(* IEC 61131-3 sources: IRIS-Project/LASAL CONTROL SOFTWARE/LasalProject_2025_09_12/Class/DiasMasterMain (part 3) *)

	push		  ecx
	push		  ebx

	L.eax		  (ebx+OneHandle.thisp)
	LZXW.ECX	(ebx+OneHandle.Address)
	push		  ecx
	push		  eax

	call		  CallUpdataRT
	add.esp		8

	pop			  ebx
	pop			  ecx

NextHandleRt
	add.ebx		sizeof (OneHandle)
	loop		  HandleLoopRt

LABEL_RtPostScan
//BLEERN START
  cmp.d     HwControl, 0
  jne       Rt_end

  call      UpdateRtPostScan_IM
//BLEERN ENDE

	jmp			  RT_end

// ****************************************************************
//  now we have to move the startpoint till we are 50usec before
// ****************************************************************

MovStartPoint

	//#SR001 Start
	L.EAX		  ud_DelayRealtime	//Time of Rt - Programm of IM
	CLR			  EDX
	L.ECX		  DmTmrResso*1000		// we have nanoseconds and we have to put in 25µs units
	DIV 		  ECX
	l.ebx		  eax
	//#SR001 End

	l.eax		  RtInterval

	sub.eax		ebx

	//#SR013 start
	cmp.b		  us_MuSecMode,1			//have we µs - Mode
	jne			  LABEL_Reserve_Std
	sub.eax		DmTimeReserveIM			//not so much reserve tim in µs - Mode
	jmp			  LABEL_EndReserve
LABEL_Reserve_Std
	//#SR013 end
	sub.eax		DmTimeReserveIM + 1		//ws005: just subtract 3 instead of ... (see above)			//#SR010 (make variable with define [instead of 3])
LABEL_EndReserve						//#SR013
  s.al		  (EDI+DmPllSyncDel)
	imul.ax		ax,DmTmrResso			//#SR009
	s.ax		  ui_RtStartPoint			//#SR009
	inc.b		  RtSSW					//ws005
	call		  LogRtSSW				//#SR008
	jmp			  RT_end

// ***********************************************************
//   read the calculated time
// ***********************************************************

ReadPoint
	clr			  eax
	l.al		  (edi+DmUserData)
	s.ax		  TimeBeforeNextSync
	inc.b		  RtSSW				//ws005
	call		  LogRtSSW			//#SR008
	jmp			  RT_end

// **********************************************************
//  now we are starting the RTProg
// **********************************************************

weAreSync
	call		  StartRealtimeProg
	inc.b		  RtSSW				//ws005
	call		  LogRtSSW			//#SR008
	jmp			  RT_end

// ***********************************************************
//   we have to wait that the PLL is locked before we start
// ***********************************************************
WaitForSync
	cmp.d		  release,16#FFFFFFFF
	je			  RT_end					// #fa 080103

	l			    (edi+DmPLLSyncState)
	test.al		DmPLLisLock
	jz			  WaitForSyncRet
	call		  StartRealtimeProg
	inc.b		  RtSSW				//ws005
	call		  LogRtSSW			//#SR008
	l.edi		  _IOSEGMENT			//#SR008
WaitForSyncRet
	L.AL		  (EDI+DmState)           // Start it always to keep the moduls alive
	OR.AL		  16#10
	S.AL		  (EDI+DmState)
	// #BS002

RT_end

	BT.W			StateCDiasSync+0,0
	JC				CDIASSyncOK
	L.EDI			CDIASSync // sync of CDIASBus
	L				  (EDI+2)
	S				  StateCDiasSync
CDIASSyncOK

	FC				WDCDIAS
RT_End1
	L.EAX	 		READY$UDINT

//#wp001
//============================ Profiler end======================================================
#ifdef  DiasMasterC_Profiler
	cmp.b 		DMC_Time_RT.initfl, 1				//schaun ob Delayzeit schon abgelaufen ist
	je			  LABEL_DMCEND
	pushad
	l.edi 		_LSL_POS
	l.edi 		( edi + DM_LSLPOS_SYSTIME )
	l.edi 		( edi + DM_LSLSYSTIME_MICROSEC )
	call		  edi								//OS_REadMicroSec - Funktion aufrufen
	s.eax 		DMC_Time_RT.stop					//Stopzeit speichern
	l.ebx 		DMC_Time_RT.start
	sub.eax		ebx								//Differenz berechnen
	sub.eax		DM_CPUconstant					//Zeit für OS_REadMicroSec - Funktion subtrahieren
	s.eax 		DMC_Time_RT.diff					//Ergebnis speicern
	l.ebx 		DMC_Time_RT.sum
	add.ebx 	eax								//Zur Summe addieren
	s.ebx 		DMC_Time_RT.sum					//Summe speichern
	l.ecx		  DMC_Time_RT.run
	inc 		  ecx								//Durchlaufzähler erhöhen
	s.ecx 		DMC_Time_RT.run					//Durchlaufzähler speichern
	cmp.eax		DMC_Time_RT._min					//mit Minimalzeit vergleichen
	jae			  LABEL_DMCcont
	s.eax 		DMC_Time_RT._min					//Minimalzeit speichern

LABEL_DMCcont
	cmp.eax 	DMC_Time_RT._max					//Mit Maximalzeit vergleichen
	jbe 		  LABEL_DMCcont1
	s.eax 		DMC_Time_RT._max					//Maximalzeit speichern

LABEL_DMCcont1
	l.eax		  ebx								//Summe in al laden
	imul.eax	eax,100							//*100 damit wir 2 Kommastellen haben
	x.edx 		edx
	idiv		  ecx								//durch Durchläufe dividieren
	s.eax		  DMC_Time_RT.avg					//Durchschnitt speichern
	popad

LABEL_DMCEND
	STI
#endif
//============================ Profiler end========================================================

END_FUNCTION
#endif

FUNCTION  DiasMasterMain::WDDIAS

	IF FirstModulFound <> 16#ff THEN	//ws005
	  IF DiasType <> 2 | RtSSw <> 4 THEN
 #IFNDEF MaxWatchdog	// #BS016
		IF ops.tAbsolute - timestamp$UDINT > 100ms | RtDebug = 1 THEN				//#SR011
			timestamp$UDINT := ops.tAbsolute;
 #ENDIF

			//**** Watchdog *************************************
			ReadKenn(FirstModulFound);

 #IFNDEF MaxWatchdog	// #BS016
		END_IF;
 #ENDIF
	  END_IF;
	END_IF;

	IF DiasType = 2 THEN
 #IFNDEF MaxWatchdog	// #BS016
		IF ops.tAbsolute - timestamp$UDINT > 100ms | RtDebug = 1 THEN				//#SR011
			timestamp$UDINT := ops.tAbsolute;
 #ENDIF

			IF (((_IOSegment$UDINT + DmControl)$^USINT)^ AND 2#10) = 0 & MasterON = 1 THEN
				MasterON := 0; // Risk is stopped => would be a watchdog
				IF Firstmodulfound <> 16#ff THEN		//ws005
          bdRTLogs.Bit6 := 1;
				END_IF;
				ImOff := 1;
			END_IF;

			//**** Watchdog for Risk (Xlinixversion 2.1) ****
			((_IOSegment$UDINT + DMWDRegister)$^USINT)^ := 1;

 #IFNDEF MaxWatchdog	// #BS016
		END_IF;
 #ENDIF
	END_IF;

END_FUNCTION

#ifdef _LSL_TARGETARCH_ARM
FUNCTION VIRTUAL GLOBAL DiasMasterMain::AddNOP
  VAR_INPUT
    RTCY		  : DINT;
    nCount		: DINT;
  END_VAR
  VAR
    i : DINT;
  END_VAR

  if (RTCY AND DmRealtime) = DmRealtime then
    ud_DelayRealtime += C_TimeNop;
  else
    ud_DelayCyclic += C_TimeNop;
  end_if;

  for i := 0 to (nCount-1) do
    (PtrCode + IPSub)^ := DbNop;

    IPSub += sizeof(RetStruct);
  end_for;

END_FUNCTION

#else
//
//	THR Aug. 21, 2003
//		Added function to add NOPs to the RISC program.  Unlike the
//		WAIT command, a NOP command CANNOT be interrupted by the
//		Cyclic Program.
//		Only for old DiasModuls
FUNCTION AWL VIRTUAL GLOBAL DiasMasterMain::AddNOP
  VAR_INPUT
    RTCY		  : DINT;
    nCount		: DINT;
  END_VAR

	l.eax		  RTCY
	and.eax		Dmrealtime

//#SR001 Start
	x.edx		  edx						//#SR003
	l.ebx		  nCount					//#SR003		//#SR009 (use ebx instead of eax register)
	imul.ebx	ebx,C_TimeNop			//#SR003		//#SR009
	CMP.EAX		Dmrealtime
	JNE			  LABEL_AN_NORT
	ADD.D		  ud_DelayRealtime,ebx	//#SR003		//#SR009
  JMP       LABEL_AN_TIMETAKEN
LABEL_AN_NORT
	ADD.D		  ud_DelayCyclic,ebx
//#SR001 End

LABEL_AN_TIMETAKEN

	call		  GetProgPointer

  l.ebx     PtrCode

	push		  ecx
	l.ecx		  nCount+0
an_loop
	l.b			  (edx+ebx),DbNop	   			// opcode NOP
	inc			  edx
	loop		  an_loop						//ws005: replaced dec,jnz with loop
	pop			  ecx

	l.eax		  RTCY
	and.eax		Dmrealtime
	call		  StoreNewPointers

END_FUNCTION
#endif

FUNCTION  DiasMasterMain::ErrorLocalSyncTrace

#ifdef HWC_LogError
  HWC_LogError(this, "@000A (DiasMasterMain::ErrorLocalSyncTrace) The constant 'NumberLocalSyncs' is defined too small !!! Remember: This is the number of maximum local Syncs !!!");
#else
	TRACE("The constant 'NumberLocalSyncs' is defined too small !!! Remember: This is the number of maximum local Syncs !!!");
#endif

END_FUNCTION

FUNCTION  DiasMasterMain::GetVerIMCIPC
  VAR_OUTPUT
    Ver(EAX)		: HDINT; // #BS016
  END_VAR
  VAR
    SigmaTekDevInfo : ^PCICONFDATA;
  END_VAR

#ifdef _LSL_TARGETARCH_X86
	SAVE_REG();
#endif

	IF pSPCIInfo <> NIL THEN
		SigmaTekDevInfo := SPCIINFO_FINDDEVICEBYNAME( "DIASIM" , 0 );
		Ver := 0;
		IF SigmaTekDevInfo <> NIL THEN
			Ver$USINT := SigmaTekDevInfo^.Version;
		END_IF;
	ELSE
		Ver := 0; // Error in OS - Interface (shouldn't be)
	END_IF;

#ifdef _LSL_TARGETARCH_X86
	RESTORE_REG();
#endif

(*
other funktions:

VAR
	pSPCIInfo     	: ^LSL_SPCIINFO;
	SigmatTekDevs	: DINT;
	SigmaTekDevInfo : ^PCICONFDATA;
	Version : USINT;
	Index : DINT;
	BaseAddress : ^VOID;
	BaseAddressLEN : UDINT;
END_VAR

	if OS_CILGET("PCICONFIG", #pSPCIInfo) then
		state:= 1;
	else
		state:= 0;
	end_if;

	// Anzahl der Einträge im InfoBlock
	SigmatTekDevs := SPCIINFO_GETDEVICECOUNT();

	for Index := 0 to SigmatTekDevs-1 do
		SigmaTekDevInfo := SPCIINFO_GETDEVICEBYINDEX( Index );
		Version := SigmaTekDevInfo^.Version;
	end_for;

	// z.B. PLL
	SigmaTekDevInfo := SPCIINFO_FINDDEVICEBYNAME( "PLL", 0 );
	SigmaTekDevInfo := SPCIINFO_FINDDEVICE( 16#0E08, 0 );
	BaseAddress := SPCIINFO_GETADDRESS( SigmaTekDevInfo );
	BaseAddressLen := SPCIINFO_GETADDRESSLEN( SigmaTekDevInfo );

	// z.B. CDIAS
	SigmaTekDevInfo := SPCIINFO_FINDDEVICEBYNAME( "CDiasBus", 0 );
	SigmaTekDevInfo := SPCIINFO_FINDDEVICE( 16#0500, 0 );
	BaseAddress := SPCIINFO_GETADDRESS( SigmaTekDevInfo );
	BaseAddressLen := SPCIINFO_GETADDRESSLEN( SigmaTekDevInfo );

*)

END_FUNCTION

FUNCTION DiasMasterMain::TraceAsyncError
	VAR_INPUT
		Place 	: UDINT;(* := 255 *)
	END_VAR
  VAR
    ptr		  : ^USINT;
    tracewd	: USINT;		// #BS012
    LogStr  : ARRAY [0..255] OF CHAR;
    NumStr  : ARRAY [0..9] OF CHAR;
  END_VAR

	if ( MasterOn <> 0 ) then		//#SR016	( because otherwise we have a lot of event messages

#ifdef _LSL_TARGETARCH_X86
		SAVE_REG();
#endif
		// #BS012 Start
		tracewd := 0;
		IF CDIASType = 2 THEN // CIPC
			IF ((CDiasI2CWatchdog+2)^ AND 1) = 1 THEN // watchdogstatus (Bit0 = 1 => watchdog)
#ifdef HWC_LogError
        HWC_LogError(this, "@0578 (DiasMasterMain::TraceAsyncError) Watchdog on CDIAS and DIAS - Bus occured !! (The RtTask of DiasMasterC - Class was set Off for more than 30ms => Hardwarereset on DIAS and CDIAS - Bus)");
#else
				// Watchdog on CDIAS and DIAS - Bus occured !! (The RtTask of DiasMasterC - Class was set Off for more than 30ms => Hardwarereset on DIAS and CDIAS - Bus)
				Trace("DiasMaster: Watchdog on CDIAS and DIAS - Bus occured !! (The RtTask of DiasMasterC - Class was set Off for more than 30ms => Hardwarereset on DIAS and CDIAS - Bus)");
				//#SR008 start
				if p_KernelLog <> NIL then
					OS_KernelLog0( "DiasMaster: Watchdog on CDIAS and DIAS - Bus occured !! (The RtTask of DiasMasterC - Class was set Off for more than 30ms => Hardwarereset on DIAS and CDIAS - Bus)" );
				end_if;
				//#SR008 end
#endif
			ELSE
				tracewd := 1;
			END_IF;
		END_IF;
		// #BS012 End
		ptr$UDINT := _IOSegment$UDINT + DMControl;
		ptr^ := 1; // Chip on risk off
		ImOff := 1;
		MasterOn := 0;
#ifdef HWC_LogError
    HWC_LogError(this, "@0582 (DiasMasterMain::TraceAsyncError) Timeout on asynchron methods !! => DiasBus is set off!!");
#else
		TRACE("DiasMaster: Timeout on asynchron methods !! => DiasBus is set off!!");
		//#SR008 start
		if p_KernelLog <> NIL then
			OS_KernelLog0( "DiasMaster: Timeout on asynchron methods !! => DiasBus is set off!!" );
		end_if;
#endif

#ifndef DIASMASTER_DISABLE_DIAS_ERROR_ON_DIRECT_ACCESS
    // if we got a place => create a dias error
    if Place <> 255 then

#ifdef HWC_LogValue1
      HWC_LogValue1(this, "@05F0 (DiasMasterMain::TraceAsyncError) Dias Error occured at place 0x{0}", Place);
#else
      _strcpy(dest:=#LogStr[0], src:="(DiasMasterMain::TraceAsyncError) Dias Error occured at place 0x");
      _itoa(udNumber:=Place, pString:=#NumStr[0]);
      _strcat(dest:=#LogStr[0], src:=#NumStr[0]);
      TRACE(#LogStr[0]);
      if p_KernelLog <> NIL then
        OS_KernelLog0(#LogStr[0]);
      end_if;
#endif

      _strcpy(dest:=#LogStr[0], src:="exec climsg 25 Dias Error occured at place 0x");
      _itoa(udNumber:=Place, pString:=#NumStr[0]);
      _strcat(dest:=#LogStr[0], src:=#NumStr[0]);

      To_OSKernel.AddToServiceProvider(command:=#LogStr[0], immediatly:=1);
    end_if;
#endif

		//#SR008 end
		// #BS012 Start
		IF tracewd THEN
#ifdef HWC_LogError
      HWC_LogError(this, "@058C (DiasMasterMain::TraceAsyncError) But no Watchdog on CDIAS and DIAS - Bus");
#else
			Trace("DiasMaster: But no Watchdog on CDIAS and DIAS - Bus");
			//#SR008 start
			if p_KernelLog <> NIL then
				OS_KernelLog0( "DiasMaster: But no Watchdog on CDIAS and DIAS - Bus" );
			end_if;
			//#SR008 end
#endif
		END_IF;
		// #BS012 End
#ifdef _LSL_TARGETARCH_X86
		RESTORE_REG();
#endif
	end_if;						//#SR016

END_FUNCTION

FUNCTION  DiasMasterMain::GetMuSec
  VAR_OUTPUT
    value(EAX)		: UDINT;
  END_VAR

#ifdef _LSL_TARGETARCH_X86
	SAVE_REG();
#endif
	value := OS_ReadMicroSec();

#ifdef _LSL_TARGETARCH_X86
	RESTORE_REG();
#endif

END_FUNCTION

#ifdef _LSL_TARGETARCH_ARM
FUNCTION VIRTUAL GLOBAL DiasMasterMain::AddRdKenn
  VAR_INPUT
    Adress		: HSINT;
    RTCY		: DINT;
    thisp		: ^void;
    callOptions 	: USINT;
  END_VAR
  VAR_OUTPUT
    Handle		: DINT;
  END_VAR

  if (RTCY AND DmRealtime) = DmRealtime then
    ud_DelayRealtime += C_TimeReadKennung;
    ui_RtDIASAccesses += 1;
  else
    ud_DelayCyclic += C_TimeReadKennung;
    ui_CyDIASAccesses += 1;
  end_if;

  (PtrCode + IPSub + RdKennStruct.Opc)^   := DbRdKenn;
  (PtrCode + IPSub + RdKennStruct.ModAdr)^ := Adress;

  ARM_EAX := RTCY$UDINT;
  ARM_EDI := thisp$UDINT;
  GetHandle(RdKennStruct.Data, callOptions);
  Handle := ARM_EAX$DINT;
  IPSub += sizeof(RdKennStruct);

END_FUNCTION

#else
// to read the identifier of a modul

FUNCTION AWL VIRTUAL GLOBAL DiasMasterMain::AddRdKenn
	VAR_INPUT
		Adress 	: HSINT;
		RTCY 	: DINT;
		thisp 	: ^void;
		callOptions 	: USINT;
	END_VAR
	VAR_OUTPUT
		Handle 	: DINT;
	END_VAR

	l.eax		  RTCY
	and.eax		Dmrealtime

//#SR001 Start
	CMP.EAX		Dmrealtime
	JNE			  LABEL_ARK_NORT
	ADD.D		  ud_DelayRealtime,C_TimeReadKennung
	inc.w		  ui_RtDIASAccesses			//#SR021
  JMP       LABEL_ARK_TIMETAKEN

LABEL_ARK_NORT
	ADD.D		  ud_DelayCyclic,C_TimeReadKennung
	inc.w		  ui_CyDIASAccesses
//#SR001 End

LABEL_ARK_TIMETAKEN

	call		  GetProgPointer

  l.ebx     PtrCode

	l.b			  (edx+ebx+RdKennStruct.Opc),DbRdKenn	   			// opcode read identifier
	l			    Adress					// adress of dias modul
	s			    (edx+ebx+RdKennStruct.ModAdr)

	l.ax		  RTCY+0
	l.edi		  thisp				    // to put into then handle

  push.b    callOptions

	push.d		RdKennStruct.Data			// direct pointer on the data
	call		  GetHandle
  add.esp   5

	s.eax		  Handle
	add.edx		sizeof (RdKennStruct)

	l.eax		  RTCY
	and.eax		Dmrealtime
	call		  StoreNewPointers

END_FUNCTION
#endif

#ifdef _LSL_TARGETARCH_ARM
FUNCTION VIRTUAL GLOBAL DiasMasterMain::AddMove
  VAR_INPUT
    RTCY		: DINT;
    thisp		: ^void;
    callOptions 	: USINT;
    SourceAddr 	: HDINT;
    DestAddr 	: HDINT;
    MoveLen 	: UDINT;
    pEnable 	: ^USINT;
    Settings 	: HDINT;
  END_VAR
  VAR_OUTPUT
    HandleMove		: DINT;
  END_VAR

  if (RTCY AND DmRealtime) = DmRealtime then
    ud_DelayRealtime += C_TimeMove;
  else
    ud_DelayCyclic += C_TimeMove;
  end_if;

  (PtrCode + IPSub + MoveStruct.Opc)^               := DbMov;
  (PtrCode$^HINT + IPSub + MoveStruct.Source)^      := (IPSub + MoveStruct.Destination)$HINT;
  (PtrCode$^HINT + IPSub + MoveStruct.Destination)^ := (IPSub + MoveStruct.Destination)$HINT;

  ARM_EAX := RTCY$UDINT;
  ARM_EDI := thisp$UDINT;
  GetHandle(MoveStruct.Source, callOptions);
  HandleMove := ARM_EAX$DINT;
  IPSub += sizeof(MoveStruct);

END_FUNCTION

#else
// BS 14.11.2001
// This command is to switch for example a bank back in im routine.
//
//[#ENGLISH]
//[<HandleMove]pointer on source (2 Byte further is destination)

FUNCTION AWL VIRTUAL GLOBAL DiasMasterMain::AddMove
	VAR_INPUT
		RTCY 	: DINT;
		thisp 	: ^void;
		callOptions 	: USINT;
		SourceAddr 	: HDINT;
		DestAddr 	: HDINT;
		MoveLen 	: UDINT;
		pEnable 	: ^USINT;
		Settings 	: HDINT;
	END_VAR
	VAR_OUTPUT
		HandleMove 	: DINT;
	END_VAR

	l.eax		  RTCY
	and.eax		Dmrealtime

//#SR001 Start
	CMP.EAX		Dmrealtime
	JNE			  LABEL_AM_NORT
	ADD.D		  ud_DelayRealtime,C_TimeMove
  JMP       LABEL_AM_TIMETAKEN

LABEL_AM_NORT
  ADD.D		  ud_DelayCyclic,C_TimeMove
//#SR001 End

LABEL_AM_TIMETAKEN

	call		  GetProgPointer

  l.ebx     PtrCode

	l.b			  (edx+ebx+MoveStruct.Opc),DbMov	   			// opcode read identifier

	L.EAX		  EDX
	ADD.EAX		MoveStruct.Destination
	S.AX		  (edx+ebx+MoveStruct.Source) // read destination
	S.AX		  (edx+ebx+MoveStruct.Destination) // save on destination

	l.ax		  RTCY+0
	l.edi		  thisp				    // to put into then handle

  push.b    callOptions

	push.d		MoveStruct.Source			// direct pointer on the data
	call		  GetHandle
  add.esp 5

	s.eax		  HandleMove
	add.edx		sizeof (MoveStruct)

	l.eax		  RTCY
	and.eax		Dmrealtime
	call		  StoreNewPointers

END_FUNCTION
#endif

FUNCTION VIRTUAL GLOBAL DiasMasterMain::GetCDiasPlaceIoSegment
  VAR_INPUT
    place		: UDINT;
  END_VAR
  VAR_OUTPUT
    IOSegment		: ^USINT;
  END_VAR

	IOSegment$UDINT :=  CDiasHwPointer$UDINT + (place*16#100)$UDINT;

END_FUNCTION

//[#ENGLISH]
//[<StateSync]0 = Busy | 1 = Sync | 2 = TimeOut
#ifdef _LSL_TARGETARCH_ARM
FUNCTION DiasMasterMain::CheckSyncModules
  VAR_INPUT
    TimeStampStart		: UDINT;
  END_VAR
  VAR_OUTPUT
    StateSync		: UDINT;
  END_VAR
  VAR
    pModule : ^WaitSyncCall;
    i : UDINT;
    MaxTime : UDINT;
  END_VAR

  // init with synchron
  StateSync := 1;

  // check if there are any sync calls
  if DiasSync.NumberCalls then
    pModule := #DiasSync.Modules[0];
    MaxTime := 0;

    // search for the max possible sync time
    for i := 0 to (DiasSync.NumberCalls - 1) do
      if (pModule^.SyncState = 0) & (pModule^.WaitTime > MaxTime) then
        MaxTime := pModule^.WaitTime;   // save the maxtime
      end_if;

      pModule += sizeof(WaitSyncCall);
    end_for;
    DiasSync.ActMaxTime := MaxTime;

    pModule := #DiasSync.Modules[0];

    // search if modules are ready
    for i := 0 to (DiasSync.NumberCalls - 1) do
      if (pModule^.SyncState = 0) then
        pModule^.SyncState := CallGetSync(thisp:=pModule^.thisp);
        if pModule^.SyncState = 0 then
          StateSync := 0;   // busy
        end_if;
      end_if;

      pModule += sizeof(WaitSyncCall);
    end_for;

    if (StateSync = 0) & ((ops.tAbsolute - TimeStampStart) > DiasSync.ActMaxTime) then
      StateSync := 2;   // timeout
    end_if;
  end_if;

END_FUNCTION
#else
FUNCTION AWL DiasMasterMain::CheckSyncModules
  VAR_INPUT
    TimeStampStart		: UDINT;
  END_VAR
  VAR_OUTPUT
    StateSync		: UDINT;
  END_VAR

// #BS014 Start
// init with synchron
	L.D			  StateSync,1

// check if there are any sync calls
	L.ECX		  DiasSync.NumberCalls
	JECXZ		  SyncReady

// search for the max possible sync time
	L.EDI		  #DiasSync.Modules[0]
	X.EAX		  EAX
SearchTime
	CMP.B		  (EDI+WaitSyncCall.SyncState),1	// if the modul is sync we cancel it
	JE			  NextObjectTime
	CMP.EAX		(EDI+WaitSyncCall.WaitTime)
	JAE			  NextObjectTime
	L.EAX		  (EDI+WaitSyncCall.WaitTime)		// save the maxtime
NextObjectTime
	ADD.EDI		SIZEOF(WaitSyncCall)
	LOOP		  SearchTime

	S.EAX		  DiasSync.ActMaxTime

// search if modules are ready
	L.EDI		  #DiasSync.Modules[0]
	L.ECX		  DiasSync.NumberCalls

SyncSearch

	CMP.B		  (EDI+WaitSyncCall.SyncState),1
	JE			  NextObject

	PUSH		  EDI
	PUSH		  ESI
	PUSH		  ECX

	X.AL		  AL

	L.EDI		  (EDI+WaitSyncCall.thisp)
	CALL		  CallGetSync

	POP			  ECX
	POP			  ESI
	POP			  EDI

	S.AL		  (EDI+WaitSyncCall.SyncState)
	CMP.AL	  1	// if sync then next obj
	JE			  NextObject
	L.D			  StateSync,0 // busy
NextObject
	ADD.EDI		SIZEOF(WaitSyncCall)
	LOOP		  SyncSearch

	CMP.D		  StateSync,1
	JE			  SyncReady

	L.EAX		  ops.tAbsolute
	SUB.EAX		TimeStampStart
	CMP.EAX		DiasSync.ActMaxTime
	JBE			  EndSyncCheck

	L.D			  StateSync,2 // timeout
	JMP			  EndSyncCheck

SyncReady

EndSyncCheck
// #BS014 End

END_FUNCTION
#endif

FUNCTION  DiasMasterMain::CallGetSync
  VAR_INPUT
    thisp(EDI)		: pHwBase;
  END_VAR
  VAR_OUTPUT
    syncchron(AL)		: USINT;
  END_VAR

	syncchron := thisp^.CheckSync();

END_FUNCTION

FUNCTION VIRTUAL GLOBAL DiasMasterMain::AddWaitSync
  VAR_INPUT
    thisp		: pVoid;
    MaxWaitTime		: UDINT;
  END_VAR

	IF DiasSync.NumberCalls * SIZEOF(WaitSyncCall) < SIZEOF(DiasSync.Modules) THEN
		DiasSync.Modules[DiasSync.NumberCalls$SINT].thisp$pVoid 	:= thisp;// #BS016
		DiasSync.Modules[DiasSync.NumberCalls$SINT].WaitTime := MaxWaitTime;// #BS016
		DiasSync.NumberCalls += 1;

		IF MaxWaitTime > DiasSync.ActMaxTime THEN
			DiasSync.ActMaxTime	:= MaxWaitTime;
		END_IF;
	ELSE

#ifdef HWC_LogError
    HWC_LogError(this, "@000B (DiasMasterMain::AddWaitSync) The constant 'MaxSyncModules' is defined too small !!!");
#else
		TRACE("The constant 'MaxSyncModules' is defined too small !!!");
#endif
	END_IF;

END_FUNCTION

FUNCTION VIRTUAL GLOBAL DiasMasterMain::Release::Read
	VAR_OUTPUT
		output (EAX) 	: HDINT;
	END_VAR

	output := Release;

END_FUNCTION

FUNCTION VIRTUAL GLOBAL DiasMasterMain::Chipstate::Read
  VAR_OUTPUT
    output		: DINT;
  END_VAR

	output := Chipstate;

END_FUNCTION

FUNCTION VIRTUAL GLOBAL DiasMasterMain::RiscState::Read
  VAR_OUTPUT
    output		: DINT;
  END_VAR

	output := RiscState;

END_FUNCTION

FUNCTION VIRTUAL GLOBAL DiasMasterMain::TimeAtRtPreEnd::Read
  VAR_OUTPUT
    output		: DINT;
  END_VAR

	output := TimeAtRtPreEnd;

END_FUNCTION

FUNCTION VIRTUAL GLOBAL DiasMasterMain::DIASRetryCounter::Read
  VAR_OUTPUT
    output		: DINT;
  END_VAR

	output := DIASRetryCounter;

END_FUNCTION

FUNCTION VIRTUAL GLOBAL DiasMasterMain::MasterON::Read
  VAR_OUTPUT
    output		: DINT;
  END_VAR

	output := MasterON;

END_FUNCTION

FUNCTION  DiasMasterMain::Risc_Off

#ifdef HWC_LogError
  HWC_LogError(this, "@0596 (DiasMasterMain::Risc_Off) RISC is set of -> DiasMasterOn = 0 and ImOff = 1");
#else
	TRACE("DiasMaster: RISC is set of -> DiasMasterOn = 0 and ImOff = 1");
	//#SR008 start
	if p_KernelLog <> NIL then
		OS_KernelLog0( "DiasMaster: RISC is set of -> DiasMasterOn = 0 and ImOff = 1" );
	end_if;
	//#SR008 end
#endif
	ImOff := 1;
	MasterOn := 0;

END_FUNCTION

#ifdef _LSL_TARGETARCH_ARM
FUNCTION VIRTUAL GLOBAL DiasMasterMain::AddIRQScan
  VAR_INPUT
    Place		: USINT;
    RTCY		: DINT;
    thisp		: ^void;
    callOptions 	: USINT;
  END_VAR
  VAR_OUTPUT
    Handle		: DINT;
  END_VAR

  if (RTCY AND DmRealtime) = DmRealtime then
    ud_DelayRealtime += C_TimeIRQScan;
  else
    ud_DelayCyclic += C_TimeIRQScan;
  end_if;

  (PtrCode + IPSub + IRQScanStruct.Opc)^    := DbIRQScan;
  (PtrCode + IPSub + IRQScanStruct.ModAdr)^ := Place;

  ARM_EAX := RTCY$UDINT;
  ARM_EDI := thisp$UDINT;
  GetHandle(IRQScanStruct.Data, callOptions);
  Handle := ARM_EAX$DINT;
  IPSub += sizeof(IRQScanStruct);

END_FUNCTION

#else
//[#ENGLISH]
//[>Place]modul number
FUNCTION AWL VIRTUAL GLOBAL DiasMasterMain::AddIRQScan
	VAR_INPUT
		Place 	: USINT;
		RTCY 	: DINT;
		thisp 	: ^void;
		callOptions 	: USINT;
	END_VAR
	VAR_OUTPUT
		Handle 	: DINT;
	END_VAR

	l.eax		  RTCY
	and.eax		Dmrealtime

	CMP.EAX		Dmrealtime
	JNE			  LABEL_AIRQ_NORT
	ADD.D		  ud_DelayRealtime,C_TimeIRQScan
  JMP       LABEL_AIRQ_TIMETAKEN

LABEL_AIRQ_NORT
	ADD.D		  ud_DelayCyclic,C_TimeIRQScan

LABEL_AIRQ_TIMETAKEN

	call		  GetProgPointer

  l.ebx     PtrCode

	l.b			  (edx+ebx+IRQScanStruct.Opc),DbIRQScan	   			// opcode IRQ identifier
	l			    Place					// place of dias modul
	s			    (edx+ebx+IRQScanStruct.ModAdr)

	l.ax		  RTCY+0
	l.edi		  thisp				    // to put into then handle

  push.b    callOptions

	push.d		IRQScanStruct.Data			// direct pointer on the data
	call		  GetHandle
  add.esp   5

	s.eax		  Handle
	add.edx		sizeof (IRQScanStruct)

	l.eax		  RTCY
	and.eax		Dmrealtime
	call		  StoreNewPointers

END_FUNCTION
#endif

#ifdef _LSL_TARGETARCH_ARM
FUNCTION VIRTUAL GLOBAL DiasMasterMain::IRQScan
  VAR_INPUT
    Place		: udint;
  END_VAR
  VAR_OUTPUT
    Data		: DINT;
  END_VAR
  VAR
    Time1, Time2  : UDINT;
    TimeoutFlag   : DINT;
  END_VAR

  if (DiasType = 2) & (ImOff = FALSE) then
#ifdef _LSL_TARGETARCH_X86
    Save_Flg();
    CLI();          // needed for async read
#endif

    Time1 := Time2 := OS_ReadMicroSec();

    while ((Time2 - Time1) <= DmConstTimeOut) do
      Time2 := OS_ReadMicroSec()
      if (_IOSegment$^USINT + DmCmdBuf1)^ AND 1 then
        exit;
      end_if;
    end_while;

    (_IOSegment$^USINT+1+DmCmdBuf1+IRQScanStruct.ModAdr)^ := Place$USINT;
    (_IOSegment$^USINT + DmCmdBuf1)^ := 0; // kill ready
    (_IOSegment$^USINT+1+DmCmdBuf1+IRQScanStruct.Opc)^ := DbIRQScan;

    Time1 := Time2 := OS_ReadMicroSec();
    TimeoutFlag := 1;

    while ((Time2 - Time1) <= DmConstTimeOut) do
      Time2 := OS_ReadMicroSec()
      if (_IOSegment$^USINT + DmCmdBuf1)^ AND 1 then
        Data := to_dint((_IOSegment$^USINT+1+DmCmdBuf1+IRQScanStruct.Data)^);
        TimeoutFlag := 0;
        exit;
      end_if;
    end_while;

    if TimeoutFlag then
      // timeout
      TraceAsyncError();
      Data := 0;
    end_if;

#ifdef _LSL_TARGETARCH_X86
    Restore_Flg();
#endif
  end_if;

END_FUNCTION

#else

FUNCTION AWL VIRTUAL GLOBAL DiasMasterMain::IRQScan
  VAR_INPUT
    Place		: udint;
  END_VAR
  VAR_OUTPUT
    Data		: DINT;
  END_VAR

  //ws005: moved to the start, since these cmp are critical
	cmp.b		  DiasType,2		//ws005
	jne			  LABEL_End		// --> it is a new Master

  CMP.B		  ImOff,1
	JE			  LABEL_End
  // /ws005

	push		  edi
	push		  ebx
	push		  eax

	L.EDI		  _IOSEGMENT

	CLR 		  EAX

 	L.ebx		  Place

	PUSHF
	CLI // needed for async read

	FC			  GetMuSec
	S.EAX		  EDX
BSyIRQ
	FC			  GetMuSec
	SUB.EAX		EDX
	TST.B		  (EDI+DmCmdBuf1),1
	JNZ			  BSyIRQConti
	CMP.EAX		DmConstTimeOut
	JA			  TimeOutError
	JMP			  BSyIRQ
BSyIRQConti

	S.Bl		  (EDI+1+DmCmdBuf1+IRQScanStruct.ModAdr)
	L.b			  (EDI+DmCmdBuf1),0		// Ready Töten
	L.B			  (EDI+1+DmCmdBuf1+IRQScanStruct.Opc),DbIRQScan

	FC			  GetMuSec
	S.EAX		  EDX
NixDaIRQ
	FC			  GetMuSec
	SUB.EAX		EDX
	TST.B		  (EDI+DmCmdBuf1),1
	JNZ			  IRQScanOkIM
	CMP.EAX		DmConstTimeOut
	JA			  TimeOutError
	JMP			  NixDaIRQ

TimeOutError
	POPF
  L.EAX     Place
  PUSH      EAX
	FC			  TraceAsyncError
  ADD.ESP   4
	L.D			  Data,0
	JMP			  LABEL_End1  //ws005

IRQScanOkIM
	LZXB.EAX	(EDI+1+DmCmdBuf1+IRQScanStruct.Data)
//	POPF				//#SR017
	S.EAX		  Data

LABEL_End1    //ws005
	POPF				//#SR017
	pop			  eax
	pop			  ebx
	pop			  edi

LABEL_End     //ws005

END_FUNCTION
#endif

//[#ENGLISH]
// This function updates the DIAS retry counter (using a function provided by the OS)
// [Globals]	_LSL_POS			:R		:OS interface structure
// [Members]	oldErrorCounter		:R/W	:calculate change
//			(S)	DiasRetryCounter	:W		:update retry counter
// [Locals]		us_actcount			:R/W	:currently read value
//				di_oldcount			:R/W	:temporary storeage of the previous value
FUNCTION DiasMasterMain::UpdateRetryCounter
  VAR
    us_actcount : usint;
    di_oldcount : dint;
    di_ret	    : dint;		//ws005
  END_VAR;

	if( pDIAS <> NIL )then	// CPU has a DIAS bus (for now only valid for CCL081)
		//ws005: consider the return value
		di_ret := OS_DIAS_ReadRegister( pDIAS, ( DIASRetryCounterOffset + 0 )$uint,  #us_actcount );
    di_oldcount := oldErrorCounter;
    oldErrorCounter := to_dint( us_actcount );
    DiasRetryCounter += oldErrorCounter - di_oldcount;
	end_if;

END_FUNCTION

//[#ENGLISH]
//Function gives back the Dias Adress, of the module which
//answer to the global sync.
FUNCTION VIRTUAL GLOBAL DiasMasterMain::GetSyncModuleNumber
  VAR_OUTPUT
    us_ModuleNr		: USINT;
  END_VAR

	us_ModuleNr := us_SyncModule;

END_FUNCTION

//[#ENGLISH]
//Function for logging Realtime steps at startup
FUNCTION  DiasMasterMain::LogRtSSW

  case RtSSW of

    1:		bdRTLogs.Bit1 := 1; //OS_KernelLog0( "DiasMaster: Pll is locked and Rt programm of intelligent master starts (1)"); 	//#SR021

    2:		bdRTLogs.Bit2 := 1; //OS_KernelLog1( "DiasMaster: We are Sync -> Rt programm of intelligent master starts again (Sync Module Place: %d) (2)", us_SyncModule ); 		//#SR021

    3:		bdRTLogs.Bit3 := 1; //OS_KernelLog2( "DiasMaster: MoveStartPointer -> Start moment of IM - programm is set (Rt - Startpoint: %dus, AddTime: %dns) (3)", ui_RtStartpoint, ui_AddTime );	//#SR021

    4:		bdRTLogs.Bit4 := 1; //OS_KernelLog1( "DiasMaster: One Time point was read -> start updating realtime tasks now (%d Rt - Dias accesses) (4)", ui_RtDIASAccesses );			//#SR021

  end_case;

END_FUNCTION

FUNCTION  DiasMasterMain::WriteRTLogs

  if bdRTLogs then
    if p_KernelLog <> NIL then
      if bdRTLogs.Bit1 then
        bdRTLogs.Bit1 := 0;
#ifdef HWC_LogError
        HWC_LogError(this, "@0514 (DiasMasterMain::WriteRTLogs) Pll is locked and Rt programm of intelligent master starts (1)");
#else
        if p_KernelLog <> NIL then
          OS_KernelLog0( "DiasMaster: Pll is locked and Rt programm of intelligent master starts (1)"); 	//#SR021
        end_if;
#endif
      end_if;
      if bdRTLogs.Bit2 then
        bdRTLogs.Bit2 := 0;
#ifdef HWC_LogValue1
        HWC_LogValue1(this, "@051E (DiasMasterMain::WriteRTLogs) We are Sync -> Rt programm of intelligent master starts again (Sync Module Place: {0}) (2)", us_SyncModule);
#else
        if p_KernelLog <> NIL then
          OS_KernelLog1( "DiasMaster: We are Sync -> Rt programm of intelligent master starts again (Sync Module Place: %d) (2)", us_SyncModule ); 		//#SR021
        end_if;
#endif
      end_if;
      if bdRTLogs.Bit3 then
        bdRTLogs.Bit3 := 0;
#ifdef HWC_LogValue2
        HWC_LogValue2(this, "@0528 (DiasMasterMain::WriteRTLogs) MoveStartPointer -> Start moment of IM - programm is set (Rt - Startpoint: {0}us, AddTime: {1}ns) (3)", ui_RtStartpoint, ui_AddTime);
#else
        if p_KernelLog <> NIL then
          OS_KernelLog2( "DiasMaster: MoveStartPointer -> Start moment of IM - programm is set (Rt - Startpoint: %dus, AddTime: %dns) (3)", ui_RtStartpoint, ui_AddTime );	//#SR021
        end_if;
#endif
      end_if;
      if bdRTLogs.Bit4 then
        bdRTLogs.Bit4 := 0;
#ifdef HWC_LogValue1
        HWC_LogValue1(this, "@0532 (DiasMasterMain::WriteRTLogs) One Time point was read -> start updating realtime tasks now (%d Rt - Dias accesses) (4)", ui_RtDIASAccesses);
#else
        if p_KernelLog <> NIL then
          OS_KernelLog1( "DiasMaster: One Time point was read -> start updating realtime tasks now (%d Rt - Dias accesses) (4)", ui_RtDIASAccesses );			//#SR021
        end_if;
#endif
      end_if;
    end_if;
  end_if;

  //Trace Message for Timesliceerror
	if us_FirstTimeSliceStart = 1 (* //#SR017 & ud_ErrorCountTimeSliceStart >= 10*) then

		us_FirstTimeSliceStart := 2;
#ifdef HWC_LogError
    HWC_LogError(this, "@05A0 (DiasMasterMain::Trace_JitterError) [SL] Rt of IM starts while Rt of DiasMaster is running!!");
#else
		trace("DiasMaster: Rt of IM starts while Rt of DiasMaster is running!!");
		if p_KernelLog <> NIL then
			OS_KernelLog0( "DiasMaster: Rt of IM starts while Rt of DiasMaster is running!!" );
		end_if;
#endif

	elsif us_FirstTimeSliceEnd = 1 (* //#SR017 & ud_ErrorCountTimeSliceEnd >= 10*) then

		us_FirstTimeSliceEnd := 2;
#ifdef HWC_LogError
    HWC_LogError(this, "@05AA (DiasMasterMain::Trace_JitterError) [SL] Timeslice overrun!!");
#else
		trace("DiasMaster: Timeslice overrun!!");
		if p_KernelLog <> NIL then
			OS_KernelLog0( "DiasMaster: Timeslice overrun!!" );
		end_if;
#endif
	end_if;

  //Watchdog Error CDIAS
  if bdRTLogs.Bit5 then
    if RTSSW <> 4 then
#ifdef HWC_LogError
      HWC_LogError(this, "@0564 (DiasMasterMain::WdCDIAS) Watchdog Error (RTSSW<>4) -> DiasMasterOn = 0 and ImOff = 1");
#else
      // Watchdog on CDIAS and DIAS - Bus occured !! (The RtTask of DiasMasterC - Class was set Off for more than 30ms => Hardwarereset on DIAS and CDIAS - Bus)
      Trace("Watchdog Error (RTSSW<>4) -> DiasMasterOn = 0 and ImOff = 1");
      //#SR008 start
      if p_KernelLog <> NIL then
        OS_KernelLog0( "Watchdog Error (RTSSW<>4) -> DiasMasterOn = 0 and ImOff = 1" );
      end_if;
      //#SR008 end
#endif
    else
#ifdef HWC_LogError
      HWC_LogError(this, "@056E (DiasMasterMain::WdCDIAS) Watchdog Error -> DiasMasterOn = 0 and ImOff = 1");
#else
      // Watchdog on CDIAS and DIAS - Bus occured !! (The RtTask of DiasMasterC - Class was set Off for more than 30ms => Hardwarereset on DIAS and CDIAS - Bus)
      Trace("Watchdog Error -> DiasMasterOn = 0 and ImOff = 1");
      //#SR008 start
      if p_KernelLog <> NIL then
        OS_KernelLog0( "Watchdog Error -> DiasMasterOn = 0 and ImOff = 1" );
      end_if;
      //#SR008 end
#endif
    end_if;
    bdRTLogs.Bit5 := 0;
  end_if;

  //Watchdog Error DIAS
  if bdRTLogs.Bit6 then

#ifdef HWC_LogError
      HWC_LogError(this, "@0009 (DiasMasterMain::WDDIAS) Watchdog on DIAS - Bus occured !! Make sure that this RtTask is called every set Real Time !! (No call for more than 130ms => Hardwarereset on DIAS - Bus)");
#else
      Trace("Watchdog on DIAS - Bus occured !! Make sure that this RtTask is called every set Real Time !! (The RtTask of DiasMasterC - Class was set Off for more than 130ms => Hardwarereset on DIAS - Bus) ");
#endif
    bdRTLogs.Bit6 := 0;
  end_if;

END_FUNCTION

//[#ENGLISH]
//For modules with old Pll (update only every ms in µs - Mode)
//[<us_update]0=no update, 1=update
FUNCTION VIRTUAL GLOBAL DiasMasterMain::GetUpdateState
  VAR_OUTPUT
    us_update		: USINT;
  END_VAR

	us_update := us_ModuleUpdate1ms;

END_FUNCTION
//[#ENGLISH]
//[<us_rt_passes]number of realtime passes before update
FUNCTION VIRTUAL GLOBAL DiasMasterMain::GetRtPasses
  VAR_OUTPUT
    us_rt_passes		: USINT;
  END_VAR

	us_rt_passes := us_RtPasses;

END_FUNCTION

//**************************************************************************
//** below this comment block are all hardware access routines which were **
//** replaced by OS calls (from version 5.44 upwards)                     **
//**    ||                                                          ||    **
//**    ||                                                          ||    **
//**   ----                                                        ----   **
//**   \  /                                                        \  /   **
//**    \/                                                          \/    **
//**************************************************************************

// /ws004
//[#ENGLISH]
// This function reads the DIAS ID of a module
// [Globals]	_IOSegment			:R
// [Members]	ImOff				:R		:master is off
//				DIAS type			:R		:intelligent <-> standard master
// [Locals]
//[>Place]		DIAS module
//[<retval]		Module ID
FUNCTION AWL DiasMasterMain::DM_DIAS_ReadKenn_x
	VAR_INPUT
    Place		: DINT;
	END_VAR
	VAR_OUTPUT
    retval		: DINT;
	END_VAR
#ifdef _LSL_TARGETARCH_X86

	L.EDI		  _IOSEGMENT

	l.al		  DiasType			//ws005
	cmp.al		2
	je			  ReadKennI			// --> intelligent
	cmp.al		1
	je			  ReadKennStd			// --> alter Master (64 k AdressRaum)

	l.eax		  16#ff				// no_kenn
	jmp			  EndReadKenn

ReadKennStd
	cmp.edi		16#d0000			// test if master in PC
	jne			  MasterFull			// no high line requiered

	l.ebx		  place
	shl.ebx		8
	add.ebx		16#ff
	pushf
	cli
	l.dx		  16#335
	l			    1
	outb
	lzxb.eax	(ebx+edi)

	push		  ax
	clr			  al
	outb
	pop			  ax

	popf
	jmp			  EndReadKenn

MasterFull
	l.ebx		  place
	shl.ebx		8
	add.ebx		16#80ff				// read kennnung
	lzxb.eax	(ebx+edi)
	jmp			  EndReadKenn

ReadKennI

// there must be some colisions with the read kennung in the OPS
	PUSHF
	CLI

// Check if someone else is working with this buffer and is not ready
	FC			  GetMuSec
	S.EAX		  EDX
BSyRdKenn
	FC			  GetMuSec				// #BS012
	TST.B		  (EDI+DmCmdBuf1),3		// #BS012
	JNZ			  RdyRdKenn
	SUB.EAX		EDX
	CMP.EAX		DmConstTimeOut
	JA			  TimeOutError
	JMP			  BSyRdKenn

RdyRdKenn

	L			    Place+0
	S  			  (EDI+1+DmCmdBuf1+Rd8Struct.ChAdr)
	l.b			  (EDI+DmCmdBuf1),0		// Ready Töten
	L.B			  (EDI+1+DmCmdBuf1+Rd8Struct.Opc),DBRdKenn
	CLR			  EAX

	FC			  GetMuSec
	S.EAX		  EDX
WaitRdKenn
	FC			  GetMuSec			// #BS012
	TST.B		  (EDI+DmCmdBuf1),3	// #BS012
	JNZ			  ReadKennRdy
	SUB.EAX		EDX
	CMP.EAX		DmConstTimeOut
	JA			  TimeOutError
	JMP			  WaitRdKenn

TimeOutError
	POPF							// #BS012
  L.EAX     255
  PUSH      EAX
	FC			  TraceAsyncError
  ADD.ESP   4
	L.EAX		  16#FF				// #BS012
	JMP			  EndReadKenn			// #BS012

ReadKennRdy
	POPF
	LZXB.EAX	(EDI+1+DmCmdBuf1+Rd8Struct.ModAdr)

EndReadKenn
	S.EAX		  retval
#endif
END_FUNCTION
//[English]
// Does a 16 Bit write access
// see Wr16Bit
FUNCTION AWL DiasMasterMain::DM_DIAS_WriteWord_x
	VAR_INPUT
		Adress 	: UDINT;
		Data 	: UINT;
	END_VAR
	VAR_OUTPUT
	state		: DINT;
	END_VAR
#ifdef _LSL_TARGETARCH_X86

  push		  edi
  push		  ebx
  push		  eax

  L.EDI		  _IOSEGMENT
  cmp.b		  DiasType,2		//ws005
  je			  Wr16IMaster		// --> it is a new Master

  // this is the old Master
  l.ebx		  Adress
  l.ax		  Data
  s.ax		  (ebx+edi+16#4000)
  jmp			  wr16ret

Wr16IMaster
  CMP.B		  ImOff,1
  JE			  Wr16Ret

  L.BX		  Adress+0

  PUSHF
  CLI	// needed for async write
  FC			  GetMuSec
  S.EAX		  EDX							// #BS012
BsyWr16
  FC			  GetMuSec
  SUB.EAX		EDX							// #BS012
  TST.B		  (EDI+DmCmdBuf1),1			// #BS012
  JNZ			  BsyWr16Conti				// #BS012
  CMP.EAX		DmConstTimeOut				// #BS012
  JA			  TimeOutError
  JMP			  BsyWr16						// #BS012
BsyWr16Conti								// #BS012

  S.BX		  (EDI+1+DmCmdBuf1+Wr16Struct.ChAdr+0)
  L.AX		  Data
  S.AX		  (EDI+1+DmCmdBuf1+Wr16Struct.Data)

  l.b			  (EDI+DmCmdBuf1),0		// Ready Töten
  L.B			  (EDI+1+DmCmdBuf1+Wr16Struct.Opc),DBWr16

  FC			  GetMuSec
  S.EAX		  EDX							// #BS012
NixDaWr16
  FC			  GetMuSec
  SUB.EAX		EDX							// #BS012
  TST.B		  (EDI+DmCmdBuf1),1			// #BS012
  JNZ			  W16OkIm						// #BS012
  CMP.EAX		DmConstTimeOut				// #BS012
  JA			  TimeOutError
  JMP			  NixDaWr16					// #BS012

TimeOutError
  POPF									// #BS012
  L.EAX     255
  PUSH      EAX
	FC			  TraceAsyncError
  ADD.ESP   4
  JMP			  wr16ret						// #BS012

W16OkIm
  POPF

wr16ret
  CLR			  EAX
  S.EAX		  State

  pop			  eax
  pop			  ebx
  pop			  edi
#endif
END_FUNCTION

//[English]
// Does a 8 Bit read access
// see Rd8Bit
FUNCTION AWL DiasMasterMain::DM_DIAS_ReadByte_x
	VAR_INPUT
		Adress 	: UDINT;
	END_VAR
	VAR_OUTPUT
    Data		: DINT;
	END_VAR
#ifdef _LSL_TARGETARCH_X86

	push		  edi
	push		  ebx
	push		  eax

	L.EDI		  _IOSEGMENT
	cmp.b		  DiasType,2		//ws005
	je			  Rd8IMaster		// --> it is a new Master

// this is the old Master
	l.ebx		  Adress
	lzxb.eax	(ebx+edi)
	s.eax		  Data
	jmp			  rd8ret

Rd8IMaster
	CLR 		  EAX
	CMP.B		  ImOff,1
	JE			  rd8Ret

 	L.BX		  Adress+0

	PUSHF
	CLI // needed for async read

	FC			  GetMuSec
	S.EAX		  EDX							// #BS012
BSyRd8
	FC			  GetMuSec
	SUB.EAX		EDX							// #BS012
	TST.B		  (EDI+DmCmdBuf1),1			// #BS012
	JNZ			  BSyRd8Conti					// #BS012
	CMP.EAX		DmConstTimeOut				// #BS012
	JA			  TimeOutError				// #BS012
	JMP			  BSyRd8						// #BS012
BSyRd8Conti									// #BS012

	S.BX		  (EDI+1+DmCmdBuf1+Rd8Struct.ChAdr+0)
	L.b			  (EDI+DmCmdBuf1),0		// Ready Töten
	L.B			  (EDI+1+DmCmdBuf1+Rd8Struct.Opc),DBRd8

	FC			  GetMuSec
	S.EAX		  EDX							// #BS012
NixDaRd8
	FC			  GetMuSec
	SUB.EAX		EDX							// #BS012
	TST.B		  (EDI+DmCmdBuf1),1			// #BS012
	JNZ			  Read8BitOkIM				// #BS012
	CMP.EAX		DmConstTimeOut				// #BS012
	JA			  TimeOutError
	JMP			  NixDaRd8					// #BS012

TimeOutError
	POPF		  							// #BS012
  L.EAX     255
  PUSH      EAX
	FC			  TraceAsyncError
  ADD.ESP   4
	L.D			  Data,0
	JMP			  rd8ret						// #BS012

Read8BitOkIM
	LZXB.EAX	(EDI+1+DmCmdBuf1+Rd8Struct.Data) // #BS012
	POPF
	S.EAX		  Data

rd8ret
	pop			  eax
	pop			  ebx
	pop			  edi
#endif
END_FUNCTION
//[English]
// Does a 16 Bit read access
// see Rd16Bit
FUNCTION AWL DiasMasterMain::DM_DIAS_ReadWord_x
	VAR_INPUT
		Adress 	: UDINT;
	END_VAR
	VAR_OUTPUT
    Data		: DINT;
  END_VAR
#ifdef _LSL_TARGETARCH_X86

	push		  edi
	push		  ebx
	push		  eax

	L.EDI		  _IOSEGMENT
	cmp.b		  DiasType,2		//ws005
	je			  Rd16IMaster		// --> it is a new Master

// this is the old Master
	l.ebx		  Adress
	lzxw.eax	(ebx+edi+16#4000)
	s.eax		  Data
	jmp			  rd16ret

Rd16IMaster
	CLR 		  EAX
	CMP.B		  ImOff,1
	JE			  rd16Ret

	L.BX		  Adress+0

	PUSHF
	CLI // needed for for async reads

	FC			  GetMuSec
	S.EAX		  EDX						// #BS012
BSyRd16
	FC			  GetMuSec
	SUB.EAX		EDX						// #BS012
	TST.B		  (EDI+DmCmdBuf1),1		// #BS012
	JNZ			  BSyRd16Conti			// #BS012
	CMP.EAX		DmConstTimeOut			// #BS012
	JA			  TimeOutError
	JMP			  BSyRd16					// #BS012
BSyRd16Conti							// #BS012

	S.BX		  (EDI+1+DmCmdBuf1+Rd8Struct.ChAdr+0)
	l.b			  (EDI+DmCmdBuf1),0		// Ready Töten
	L.B			  (EDI+1+DmCmdBuf1+Rd8Struct.Opc),DBRd16

	FC			  GetMuSec
	S.EAX		  EDX						// #BS012
NixDaRd16
	FC			  GetMuSec
	SUB.EAX		EDX						// #BS012
	TST.B		  (EDI+DmCmdBuf1),1		// #BS012
	JNZ			  Read16BitOKIM			// #BS012
	CMP.EAX		DmConstTimeOut			// #BS012
	JA			  TimeOutError
	JMP			  NixDaRd16				// #BS012

TimeOutError
	POPF								// #BS012
  L.EAX     255
  PUSH      EAX
	FC			  TraceAsyncError
  ADD.ESP   4
	L.D			  Data,0
	JMP			  rd16ret

Read16BitOKIM
	LZXW.EAX	(EDI+1+DmCmdBuf1+Rd8Struct.Data+0)	// #BS012
	POPF
	S.EAX		  Data

rd16ret
	pop			  eax
	pop			  ebx
	pop			  edi
#endif
END_FUNCTION
//[English]
// Does a 8 Bit write access (control area)
// see WrCntr
FUNCTION AWL DiasMasterMain::DM_DIAS_WriteCtrl_x
	VAR_INPUT
    adress		: DINT;
		Data 	: USINT;
	END_VAR
	VAR_OUTPUT
    state		: DINT;
	END_VAR
#ifdef _LSL_TARGETARCH_X86

	push		  edi
	push		  ebx
	push		  eax

	L.EDI		  _IOSEGMENT
	cmp.b		  DiasType,2			//ws005
	je			  WrCntrIMaster		// --> it is a new Master

	CMP.EDI		16#D0000
	JNE			  StdMasterCPU

	PUSH		  DX
	PUSHF
	CLI

	l.dx		  16#335
	l			    1
	outb // switch controller

	l.ebx		  Adress
	l.al		  Data
	s.al		  (ebx+edi)

	clr			  al
	outb // switch controller back

	POPF
	POP			  DX
	jmp			  WrCntrRet

// this is the old Master
StdMasterCPU
	l.ebx		  Adress
	l.al		  Data
	s.al		  (ebx+edi+16#8000)
	jmp			  WrCntrRet

WrCntrIMaster
	L.BX		  Adress+0

	CMP.B		  ImOff,1
	JE			  WrCntrRet

	PUSHF
	CLI			// needed for async access

	FC			  GetMuSec
	S.EAX		  EDX							// #BS012
BsyCntw
	FC			  GetMuSec
	SUB.EAX		EDX							// #BS012
	TST.B		  (EDI+DmCmdBuf1),1			// #BS012
	JNZ			  BSyCntwConti				// #BS012
	CMP.EAX		DmConstTimeOut				// #BS012
	JA			  TimeOutError
	JMP			  BsyCntw						// #BS012
BSyCntwConti								// #BS012

	S.BX		  (EDI+1+DmCmdBuf1+CntrlStruct.chAdr+0)
	L		      Data
	S			    (EDI+1+DmCmdBuf1+CntrlStruct.Data)
	l.b			  (EDI+DmCmdBuf1),0		// Ready Töten
	L.B			  (EDI+1+DmCmdBuf1+CntrlStruct.OPC),DbCntrl

	FC			  GetMuSec
	S.EAX		  EDX							// #BS012
NixDaCnt
	FC			  GetMuSec
	SUB.EAX		EDX							// #BS012
	TST.B		  (EDI+DmCmdBuf1),1			// #BS012
	JNZ			  WrCntrOK					// #BS012
	CMP.EAX		DmConstTimeOut				// #BS012
	JA			  TimeOutError
	JMP			  NixDaCnt					// #BS012

TimeOutError
	POPF
  L.EAX     255
  PUSH      EAX
	FC			  TraceAsyncError
  ADD.ESP   4
	JMP			  WrCntrRet

WrCntrOK
	POPF

WrCntrRet
	clr			  eax
	S.EAX		  State

	pop 		  eax
	pop 		  ebx
	pop 		  edi
#endif
END_FUNCTION
//[English]
// Does a 8 Bit write access
// see Wr8Bit
FUNCTION AWL DiasMasterMain::DM_DIAS_WriteByte_x
	VAR_INPUT
		Adress 	: UDINT;
		Data 	: USINT;
	END_VAR
	VAR_OUTPUT
    State		: DINT;
	END_VAR
#ifdef _LSL_TARGETARCH_X86

	push		  edi
	push		  ebx
	push		  eax

	L.EDI		  _IOSEGMENT
	cmp.b		  DiasType,2		//ws005
	je			  Wr8IMaster		// --> it is a new Master

// this is the old Master
	l.ebx		  Adress
	l.al		  Data
	s.al		  (ebx+edi)
	jmp			  wr8ret

Wr8IMaster

	CMP.B		  ImOff,1
	JE			  Wr8Ret

	L.BX		  Adress+0

	PUSHF
	CLI // needed for async write
	FC			  GetMuSec
	S.EAX		  EDX					// #BS012
BsyWr8
	FC			  GetMuSec
	SUB.EAX		EDX					// #BS012
	TST.B		  (EDI+DmCmdBuf1),1	// #BS012
	JNZ			  BSyWr8Conti			// #BS012
	CMP.EAX		DmConstTimeOut		// #BS012
	JA			  TimeOutError
	JMP			  BsyWr8				// #BS012
BSyWr8Conti

	S.BX		  (EDI+1+DmCmdBuf1+Wr8Struct.ChAdr+0)
	L		      Data
	S			    (EDI+1+DmCmdBuf1+Wr8Struct.Data+0)

	l.b			  (EDI+DmCmdBuf1),0		// Ready Töten
	L.B			  (EDI+1+DmCmdBuf1+Wr8Struct.Opc),DBWr8

	FC			  GetMuSec
	S.EAX		  EDX
NixDaWr8
	FC			  GetMuSec
	SUB.EAX		EDX					// #BS012
	TST.B		  (EDI+DmCmdBuf1),1	// #BS012
	JNZ			  W8OkIm				// #BS012
	CMP.EAX		DmConstTimeOut		// #BS012
	JA			  TimeOutError		// #BS012
	JMP			  NixDaWr8			// #BS012

TimeOutError
	POPF							// #BS012
  L.EAX     255
  PUSH      EAX
	FC			  TraceAsyncError
  ADD.ESP   4
	JMP			  Wr8Ret				// #BS012

W8OkIm
	POPF

Wr8Ret
	CLR			  EAX
	S.EAX		  State
	pop			  eax
	pop			  ebx
	pop			  edi
#endif
END_FUNCTION

FUNCTION  DiasMasterMain::CCLWatchdog_Trigger

	OS_WATCHDOG_TRIGGER();

END_FUNCTION

#ifdef _LSL_TARGETARCH_ARM
FUNCTION DiasMasterMain::SendSync

  if p_NewPll = 0 then
    if CDIASSync then
      if us_MuSecMode then                //is µs Mode active ?
        us_ModuleUpdate1ms := (CDIASSync + 3)^ AND 1; //we need only Bit0

        if us_RtPasses = us_Counter_us then   //can we send sync signal (every ms in µs - Mode) ?
          us_Counter_us := 1;
          (CDIASSync)^ := 0;
          if DiasType = 2 then
            (_IOSegment$^USINT+DmPllSyncAdr)^ := 0;
          end_if;
        else
          us_Counter_us += 1;
        end_if;
      else
        us_Counter_us := 1;
        (CDIASSync)^ := 0;                // sync of CDIASBus
        if DiasType = 2 then
          (_IOSegment$^USINT+DmPllSyncAdr)^ := 0;
        end_if;
      end_if;
    else
      if DiasType = 2 then
        (_IOSegment$^USINT+DmPllSyncAdr)^ := 0;
      end_if;
    end_if;
  end_if;

END_FUNCTION
#else
FUNCTION AWL DiasMasterMain::SendSync			//#SR014

	cmp.d			  p_NewPll, 0					//#SR016
	jne				  LABEL_EndPllSync			//#SR016

	cmp.d     	CDIASSync,0					//#SR014
	je        	LABEL_SendDiasSync			//#SR014

	//#SR013 start
	cmp.b			  us_MuSecMode,1						//is µs Mode active
	jne				  LABEL_PllSync

	l.b				  us_ModuleUpdate1ms,0				//do not update (for modules with old Pll)
	l.edi			  CDIASSync
	l.al			  ( edi + 3 )							//check sync register (Bit0 = Sync Out)
	and.al			1									//we need only Bit0
	o.al			  al									//is bit set
	jz				  LABEL_NoSyncRead
	l.b				  us_ModuleUpdate1ms,1				//modules can update (for modules with old pll)

LABEL_NoSyncRead
 	l.edi			  _IOSegment
	l.al			  us_RtPasses
 	cmp.al			us_Counter_us						//can we send sync signal (every ms in µs - Mode)
	je				  LABEL_PllSync
	inc.b			  us_Counter_us						//increment counter
	jmp				  LABEL_EndPllSync

LABEL_PllSync
	l.b				  us_Counter_us,1
	//#SR013 end

  L.EDI			  CDIASSync // sync of CDIASBus
	S				    (EDI)

	//#SR014 start
LABEL_SendDiasSync
	cmp.b			  DiasType,2
	jne				  LABEL_EndPllSync
	//#SR014 end

	L.EDI			  _IOSEGMENT
//--- Sync To Master PLL --
	S				    (EDI+DmPllSyncAdr)
LABEL_EndPllSync

END_FUNCTION
#endif

FUNCTION DiasMasterMain::FinishIMProg
  VAR
    i		   : UDINT;
  END_VAR

	if DiasType = 2  then  // test if we have a IMaster
		if release <> 16#ffffffff then  // #fa 080103

			//#SR005 Start
			p_ModuleRetryCnt := ( _IOSegment$UDINT + 16#F200 )$^ModuleRetryCnt;
			for i := 0 to 63 do
				( ( p_ModuleRetryCnt + i )$^USINT )^ := 0;
			end_for;
			//#SR005 End

			//#SR021 start
			//add Realtime Time offset for IM (actually for CIC012)
			ud_DelayRealtime += ( ui_AddTime * ui_RtDIASAccesses );
      ud_DelayCyclic += ( ui_AddTime * ui_CyDIASAccesses );
			//#SR021 end

			//#SR004 Start
			if IPMainCy > ( ud_IMMemory / 4 )$DINT then//DmCallRes * sizeof( CallStruct ) then
#ifdef HWC_LogError
        HWC_LogError(this, "@05B4 (DiasMasterMain::FinishIMProg) Too many cyclic calls");
#else
				TRACE("DiasMaster: Too many cyclic calls");
				//#SR008 start
				if p_KernelLog <> NIL then
					OS_KernelLog0( "DiasMaster: Too many cyclic calls");
				end_if;
				//#SR008 end
#endif
				MasterOn := 0;
				ImOff := 1;

			elsif IPMainRt >  ( ud_IMMemory / 4 )$DINT then//DmCallRes * sizeof( CallStruct ) then
#ifdef HWC_LogError
        HWC_LogError(this, "@05BE (DiasMasterMain::FinishIMProg) Too many realtime calls");
#else
        TRACE("DiasMaster: Too many realtime calls");
				//#SR008 start
				if p_KernelLog <> NIL then
					OS_KernelLog0( "DiasMaster: Too many realtime calls");
				end_if;
				//#SR008 end
#endif
				MasterOn := 0;
				ImOff := 1;

      elsif IPSub > ( ud_IMMemory / 2 )$DINT then
#ifdef HWC_LogError
        HWC_LogError(this, "@000C (DiasMasterMain::FinishIMProg) Program of intelligent master is too large");
#else
        TRACE("DiasMaster: Program of intelligent master is too large");
				//#SR008 start
				if p_KernelLog <> NIL then
					OS_KernelLog0( "DiasMaster: Program of intelligent master is too large");
				end_if;
				//#SR008 end
#endif
				MasterOn := 0;
				ImOff := 1;

      else
	  		//#SR004 End

				//#SR015 start
				//calculate Rt - Startpoint (detailed description see Methode "RtWorkCIPC" Label "MovestartPoint"
				if ( us_MusecMode ) then
					( ( _IOSegment$UDINT + DmPllSyncDel )$^USINT )^ := ( RtInterval$UDINT - ( ud_DelayRealtime / ( DmTmrResso * 1000 ) ) - DmTimeReserveIM )$USINT;
				else
					( ( _IOSegment$UDINT + DmPllSyncDel )$^USINT )^ := ( RtInterval$UDINT - ( ud_DelayRealtime / ( DmTmrResso * 1000 ) ) - DmTimeReserveIM - 1 )$USINT;
				end_if;
				//#SR015 end

				LinkMaster();
				LoadCyclicProg();
				LoadRealtimeProg();
        LoadRtCyCode();
				StartCyclicProg();
				DIASRetryCounter :=0;
			end_if;	//#SR004

			#ifndef OldDiasXilinx										//#SR013
				//we have to set the pointer for RTBSync Realtimeprog

      HandlesRT[0].thisp := ( SyncCall.Read() )$^HwBase;    //===HF
			#endif

      RtTimeIM_us := ud_DelayRealtime/1000;
      CyTimeIM_us := ud_DelayCyclic/1000;

			//#SR013 start
			if _RtOSversion >= 16#1132 & us_MuSecMode then
				if ud_DelayRealtime > ui_ClockTicks * 1000 / 2 then
#ifdef HWC_LogError
          HWC_LogError(this, "@05D2 (DiasMasterMain::FinishIMProg) Time of realtime - program of intelligent master is to long. Diasbus is set off");
#else
					TRACE("Time of realtime - program of intelligent master is to long. Diasbus is set off");
#endif
					MasterOn := 0;
					ImOff := 1;
				elsif (ud_DelayRealtime + ud_DelayCyclic) > ui_ClockTicks * 1000 / 2 then
#ifdef HWC_LogError
          HWC_LogError(this, "@05C8 (DiasMasterMain::FinishIMProg) Warning: Cyclic - program of intelligent master can't be done in 1 run");
#else
					TRACE("Warning: Cyclic - program of intelligent master can't be done in 1 run");
#endif
        end_if;
      else
				if ud_DelayRealtime > (sd_PllTimeGlob_us$UDINT * 1000) then
#ifdef HWC_LogError
          HWC_LogError(this, "@05D2 (DiasMasterMain::FinishIMProg) Time of realtime - program of intelligent master is to long. Diasbus is set off");
#else
					TRACE("Time of realtime - program of intelligent master is to long. Diasbus is set off");
#endif
					MasterOn := 0;
					ImOff := 1;
				elsif (ud_DelayRealtime + ud_DelayCyclic) > (sd_PllTimeGlob_us$UDINT * 1000) then
#ifdef HWC_LogError
          HWC_LogError(this, "@05C8 (DiasMasterMain::FinishIMProg) Warning: Cyclic - program of intelligent master can't be done in 1 run");
#else
					TRACE("Warning: Cyclic - program of intelligent master can't be done in 1 run");
#endif
        end_if;
			end_if;
			//#SR013 end
		end_if;

 		IF CDiasType = 2 THEN
      this^.control.pmeth^.rtwork := #RtWorkIMCIPC();
      CorrectMyTaskTime();
 		END_IF;
	else

 		this^.control.pmeth^.cywork :=#CyWorkStdMas();

 		if _IOSegment <> 16#d0000 then
      // we overload our rtwork and cywork funktion
      // because we have a standard master
      this^.control.pmeth^.rtwork :=#RtWorkStdMas();
      rtssw :=4;	// it is standard so no setup phase
 		else
      this^.control.pmeth^.rtwork :=#RtWorkStdMasIPC();
      rtssw :=4;	// it is standard so no setup phase
 		end_if;

	end_if;

	//#SR016 start
	if ( p_NewPll <> NIL ) & (DiasType = 2) then
		this^.control.pmeth^.rtwork :=#RtWorkETV();
	end_if;
	//#SR016 end

  if ImOff then
#ifdef HWC_LogError
    HWC_LogError(this, "@05DC (DiasMasterMain::FinishIMProg) Intelligent master has been switched off");
#else
    //#SR008 start
    if p_KernelLog <> NIL then
      OS_KernelLog0( "DiasMaster: Intelligent master has been switched off" );
    end_if;
    //#SR008 end
#endif
  end_if;

END_FUNCTION

FUNCTION DiasMasterMain::LastInit
  VAR
    ActualTime  : UDINT;
    ErrorSync   : USINT;	// #BS011
    StateSync   : UDINT; // #BS011
    i		        : UDINT;
    ptrS	      : ^WaitSyncCall;
    sz_name	    : ARRAY[ 0..255 ] OF CHAR;	//ws006
  END_VAR

	IF _LSL_POS^.piTask^$MYLSL_ITASK.SetNbrOfLdrPhaseObjects <> NIL
 		& _LSL_POS^.piTask^$MYLSL_ITASK.MoveObject THEN// nur wenn funktionen verfügbar

		// ****** first synchronize the IM ****************************************
 		// bring me to the first position
 		if ( HwControl = 0 ) then			//#SR014

			OS_MoveObject(this,2,1);
 			OS_SetNbrOfLdrPhaseObjects(1);
		end_if;												//#SR014

 		// now wait max 1 sek to get sync otherwise start APL and give
 		// error message to develloper
 		ActualTime := ops.tAbsolute;
 		ErrorSync  := 0; // #BS011

	 	// now we wait till the Master is synchron
 		while ((ops.tAbsolute - ActualTime) < 5secs) do
      if rtssw = 4 then
        cywork();
      end_if;
      if (CyclicReady AND 1) & (RealtimeReady AND 1) then
#ifdef HWC_LogError
        HWC_LogError(this, "@053C (DiasMasterMain::LastInit) Init ends");
#else
        //#SR008 start
        if p_KernelLog <> NIL then
          OS_KernelLog0( "DiasMaster: Init ends" );
        end_if;
        //#SR008 end
#endif
        EXIT;	// --> READY start
      end_if;
 		end_while;

 		if ((ops.tAbsolute - ActualTime) >= 5secs) then
#ifdef HWC_LogError
      HWC_LogError(this, "@05E6 (DiasMasterMain::LastInit) Timeout while synchronization. DIAS Master is not ready (startup fault)!");
#else
      TRACE("DiasMaster: Timeout while synchronization. DIAS Master is not ready (startup fault)!");
			//#SR008 start
			if p_KernelLog <> NIL then
				OS_KernelLog0( "DiasMaster: Timeout while synchronization. DIAS Master is not ready (startup fault)!");
			end_if;
			//#SR008 end
#endif
      ErrorSync := 1;
 		end_if;
	end_if;

		// ****** then synchronize all DiasModules if necessary ***********************
	// #BS011
	IF WaitSync & ErrorSync = 0 THEN
		ActualTime := ops.tAbsolute;
		StateSync := CheckSyncModules(ActualTime);
		WHILE StateSync = 0 DO
			cywork();
			StateSync := CheckSyncModules(ActualTime);
		END_WHILE;
		IF StateSync = 2 THEN
			// on timeout we trace the objectnames
			IF DiasSync.NumberCalls THEN
				ptrS := #DiasSync.Modules[0];
#ifdef HWC_LogError
        HWC_LogError(this, "@000D (DiasMasterMain::LastInit) Timeout on synchronizing modules on objects:");
#else
				Trace("Timeout on synchronizing modules on objects:");
#endif
				FOR i := 0 TO DiasSync.NumberCalls-1 DO
					IF PtrS^.SyncState = 0 THEN
						IF PtrS^.thisp <> NIL THEN
							//ws006
							_GetObjName( PtrS^.thisp$^VirtualBase, #sz_name[ 0 ] );
#ifdef HWC_LogError
              HWC_LogError(this, #sz_name[ 0 ]);
#else
							trace( #sz_name[ 0 ] );
#endif
						ELSE
#ifdef HWC_LogError
              HWC_LogError(this, "Object with NIL Pointer !!");
#else
							Trace("Object with NIL Pointer !!");
#endif
						END_IF;
					END_IF;
					PtrS += SIZEOF(WaitSyncCall);
				END_FOR;
			END_IF;
		END_IF;
	END_IF;
	// #BS011

END_FUNCTION

#ifdef _LSL_TARGETARCH_ARM
FUNCTION VIRTUAL GLOBAL DiasMasterMain::RtWorkETV
  VAR_INPUT
    EAX		: UDINT;
  END_VAR
  VAR_OUTPUT
    state		: UDINT;
  END_VAR
  VAR
    Temp      : DINT;
    pHandle   : ^OneHandle;
    i         : UDINT;
  //-------------------------------------Profiler Start----------------------------------------------
  #ifdef DiasMasterC_Profiler
    MuSecTime : UDINT;
  END_VAR

  MuSecTime := OS_ReadMicroSec();
  //Anfangsdelay abwarten
	if MuSecTime - DMC_Time_RT.init > DM_ProfilerDelay then
    DMC_Time_RT.start  := MuSecTime;    //Startzeit nehmen
    DMC_Time_RT.initfl := FALSE;        //Initflag löschen
  else
    DMC_Time_RT.initfl := TRUE;         //Initflag setzen
  end_if;
//-------------------------------------Profiler End------------------------------------------------
#else
  END_VAR
#endif

  if b_PllInit = FALSE then
    StartPll();
    b_PllInit := TRUE;
  end_if;

  if (ImOff = FALSE) then
    //look if Rt program of IM is finished
    if (ops.SysState = C_RUNRAM) & (_IOSegment$^USINT + DmUserData + 3)^ then
      ud_ErrorCountTimeSliceEnd += 1;
      if us_FirstTimeSliceEnd = 0 then
        us_FirstTimeSliceEnd := 1;
      end_if;
    end_if;

    //Reset Byte to find out if Rt of IM starts while Rt of DM is running
    (_IOSegment$^USINT + DmUserData + 4)^ := 0;

    case RtSSW of

        // ***********************************************************
        //   we have to wait that the PLL is locked before we start
        // ***********************************************************
      0:

        if Release <> 16#FFFFFFFF then
          StartRealtimeProg();
          RtSSW += 1;
          LogRtSSW();
        end_if;

        // **********************************************************
        //  now we are starting the RTProg
        // **********************************************************
      1:

        StartRealtimeProg();
        RtSSW += 1;
        LogRtSSW();

        // ****************************************************************
        //  now we have to move the startpoint till we are 50usec before
        // ****************************************************************
      2:

        if us_MuSecMode then
          Temp := RtInterval - (ud_DelayRealtime / (DmTmrResso * 1000))$DINT - DmTimeReserveIM;
        else
          Temp := RtInterval - (ud_DelayRealtime / (DmTmrResso * 1000))$DINT - (DmTimeReserveIM + 1);
        end_if;
        (_IOSegment$^USINT + DmPllSyncDel)^ := Temp$USINT;
        ui_RtStartPoint := Temp$UINT * DmTmrResso;
        RtSSW += 1;
        LogRtSSW();

        // ***********************************************************
        //   read the calculated time
        // ***********************************************************
      3:

        TimeBeforeNextSync := to_uint((_IOSegment$^USINT + DmUserData)^);
        RtSSW += 1;
        LogRtSSW();

        // ***************************************************************
        //   do the refresh of I/O
        // ***************************************************************
      4:

        // get rtload of im
        TimeAtRtPreEnd := (_IOSegment$^USINT + DmUserData)^ * DmTmrResso;
        Rt_Load := ((TimeAtRtPreEnd - ui_RtStartPoint) * 1000) / sd_PllTimeGlob_us;

        RealtimeReady := TRUE;

        // now take data and call update methods with thispointer
        if HandleNrRT then
          pHandle := #HandlesRT[0];
          for i := 0 to HandleNrRT-1 do
            if pHandle^.Typ AND DmCallProg then
              pHandle^.thisp^.UpdateRt(pHandle^.Address);
            end_if;

            pHandle += sizeof(OneHandle);
          end_for;

          if HwControl = 0 then
            UpdateRtPostScan_IM();
          end_if;
        end_if;
    end_case;

    if (StateCDiasSync AND 1) = 0 then
      StateCDiasSync := (CDIASSync + 2)^;
    end_if;

    WDDIAS();
  end_if;

  state := READY;

//-------------------------------------Profiler Start----------------------------------------------
#ifdef DiasMasterC_Profiler
  //schaun ob Delayzeit schon abgelaufen ist
  if DMC_Time_RT.initfl = FALSE then
    MuSecTime := OS_ReadMicroSec();

    DMC_Time_RT.stop := MuSecTime;        //Stopzeit speichern

    MuSecTime -= DMC_Time_RT.start;       //Differenz berechnen
    MuSecTime -= DM_CPUconstant;          //Zeit für OS_REadMicroSec - Funktion subtrahieren

    DMC_Time_RT.diff := MuSecTime;        //korr. Differenz speichern
    DMC_Time_RT.sum  += MuSecTime;        //Zur Summe addieren

    DMC_Time_RT.run  += 1;                //Durchlaufzähler erhöhen

    if MuSecTime < DMC_Time_RT._min then
      DMC_Time_RT._min := MuSecTime;      //Minimalzeit speichern
    end_if;

    if MuSecTime > DMC_Time_RT._max then
      DMC_Time_RT._max := MuSecTime;      //Maximalzeit speichern
    end_if;

    //Durchschnitt berechnen
    //*100 damit wir 2 Kommastellen haben
    DMC_Time_RT.avg := DMC_Time_RT.sum * 100 / DMC_Time_RT.run;
  end_if;

#endif
//-------------------------------------Profiler End------------------------------------------------
END_FUNCTION
#else
FUNCTION AWL VIRTUAL GLOBAL DiasMasterMain::RtWorkETV				//#SR016
  VAR_INPUT
    EAX		: UDINT;
  END_VAR
  VAR_OUTPUT
    state		: UDINT;
  END_VAR

//#wp001
//============================ Profiler start======================================================
#ifdef  DiasMasterC_Profiler
	CLI											//damit keine Interrupts die Messung stören
	push 		  edi
	push 		  eax
	l.edi 		_LSL_POS
	l.edi 		( edi + DM_LSLPOS_SYSTIME )
	l.edi 		( edi + DM_LSLSYSTIME_MICROSEC )
	call		  edi								//OS_ReadMicroSec - Funktion aufrufen
	l.ebx		  eax
	sub.ebx		DMC_Time_RT.init					//Anfangsdelay abwarten
	cmp.ebx		DM_ProfilerDelay
	jle			  LABEL_DMCPREEND
	s.eax 		DMC_Time_RT.start					//Startzeit nehmen
	x.cl		  cl
	s.cl		  DMC_Time_RT.initfl				//Initflag löschen
	jmp 		  LABEL_DMCstartfunc

LABEL_DMCPREEND
	l.b		    DMC_Time_RT.initfl,1					//Initflag setzen

LABEL_DMCstartfunc
	pop 		  eax
	pop 		  edi
#endif
//============================ Profiler end========================================================

	//#SR022 start
	cmp.b			b_PllInit, TRUE
	je				LABEL_NoStart

	//in first run we start pll
	call			StartPll
	l.b				b_PllInit, TRUE
LABEL_NoStart
	//#SR022 end

	CMP.B			ImOff,1
	JE				RT_End1

	cmp.w			ops.SysState,1					//look if CPU is in RunRam
	jne				LABEL_Continue

  	l.edi			_IOSegment
	l.bl			( edi + DmUserData + 3 )		//look if Rt program of IM is finished
	o.bl			bl
	jz				LABEL_Continue
	inc.d			ud_ErrorCountTimeSliceEnd
	cmp.b			us_FirstTimeSliceEnd,0
	jne				LABEL_Continue

	l.b				us_FirstTimeSliceEnd,1
LABEL_Continue
  l.edi			_IOSegment
	l.b				( edi + DmUserData + 4 ), 0		//Reset Byte to find out if Rt of IM starts while Rt of DM is running

	lzxb.eax	RtSSW
	shl.eax		3           //save some time here
	add.eax		#RtSel
	jmp			  eax

RtSel
	jmp			WaitForSync			// 0 : wait till PLL in locked
	rcl.eax 	0					//ws005: simple placeholder (does really nothing)
	jmp			weAreSync			// 1 : wait one period to get a right time
	rcl.eax 	0					//ws005: simple placeholder (does really nothing)
	jmp			MovStartPoint		// 2 : mov start point to the right pos
	rcl.eax 	0					//ws005: simple placeholder (does really nothing)
	jmp			readpoint           // 3 : read one time the point
	rcl.eax 	0					//ws005: simple placeholder (does really nothing)
	jmp			RtRefresh			// 4 : do the realtime refresh

// ***************************************************************
//   do the refresh of I/O
// ***************************************************************

RtRefresh

// *************************************************
//  read the time point
// *************************************************
	lzxb.eax	(edi+DmUserData)
	imul.ax		ax,DmTmrResso
	s.eax 		TimeAtRtPreEnd

	//***********calculate Rt - usage rate***********************
	lzxw.ebx	ui_RtStartPoint
	sub.eax		ebx
	imul.eax	eax,1000
	x.edx		  edx
	l.ebx		  sd_PllTimeGlob_us
	div			  ebx
	s.eax		  Rt_Load

// **************************************************
//  now take data and call update function with thisp
// **************************************************
	l.b			  RealtimeReady,1

	l.ebx		  #HandlesRt
	lzxw.ecx	HandleNrRt
	jecxz		  LABEL_RtPostScan

HandleLoopRt
	test.w		(ebx+OneHandle.Typ),DmCallProg
	jz			  NextHandleRt

	push		  ecx
	push		  ebx

	L.eax		  (ebx+OneHandle.thisp)
	LZXW.ECX	(ebx+OneHandle.Address)
	push		  ecx
	push		  eax

	call		  CallUpdataRT
	add.esp		8

	pop			  ebx
	pop			  ecx

NextHandleRt
	add.ebx		sizeof (OneHandle)
	loop		  HandleLoopRt

LABEL_RtPostScan
//BLEERN START
  cmp.d     HwControl, 0
  jne       Rt_end

  call      UpdateRtPostScan_IM
//BLEERN ENDE

	jmp			  RT_end

// ****************************************************************
//  now we have to move the startpoint till we are 50usec before
// ****************************************************************

MovStartPoint
	L.EAX		  ud_DelayRealtime	//Time of Rt - Programm of IM
	CLR			  EDX
	L.ECX		  DmTmrResso*1000		// we have nanoseconds and we have to put in 25µs units
	DIV 		  ECX
	l.ebx		  eax

	l.eax		  RtInterval
	sub.eax		ebx
	cmp.b		  us_MuSecMode,1			//have we µs - Mode
	jne			  LABEL_Reserve_Std
	sub.eax		DmTimeReserveIM			//not so much reserve tim in µs - Mode
	jmp			  LABEL_EndReserve
LABEL_Reserve_Std
	sub.eax		DmTimeReserveIM + 1
LABEL_EndReserve
	s.al		  (EDI+DmPllSyncDel)
	imul.ax		ax,DmTmrResso
	s.ax		  ui_RtStartPoint
	inc.b		  RtSSW
	call		  LogRtSSW
	jmp			  RT_end

// ***********************************************************
//   read the calculated time
// ***********************************************************

ReadPoint
	clr			  eax
	l.al		  (edi+DmUserData)
	s.ax		  TimeBeforeNextSync
	inc.b		  RtSSW
	call		  LogRtSSW
	jmp			  RT_end

// **********************************************************
//  now we are starting the RTProg
// **********************************************************

weAreSync
	call		  StartRealtimeProg
	inc.b		  RtSSW
	call		  LogRtSSW
	jmp			  RT_end

// ***********************************************************
//   we have to wait that the PLL is locked before we start
// ***********************************************************
WaitForSync
	cmp.d		  release,16#FFFFFFFF
	je			  RT_end

	call		  StartRealtimeProg
	inc.b		  RtSSW
	call		  LogRtSSW
RT_end

	FC				WDCDIAS
RT_End1
	L.EAX	 		READY$UDINT

//#wp001
//============================ Profiler end======================================================
#ifdef  DiasMasterC_Profiler
	cmp.b 		DMC_Time_RT.initfl, 1				//schaun ob Delayzeit schon abgelaufen ist
	je			LABEL_DMCEND
	pushad
	l.edi 		_LSL_POS
	l.edi 		( edi + DM_LSLPOS_SYSTIME )
	l.edi 		( edi + DM_LSLSYSTIME_MICROSEC )
	call		  edi								//OS_REadMicroSec - Funktion aufrufen
	s.eax 		DMC_Time_RT.stop					//Stopzeit speichern
	l.ebx 		DMC_Time_RT.start
	sub.eax		ebx								//Differenz berechnen
	sub.eax		DM_CPUconstant					//Zeit für OS_REadMicroSec - Funktion subtrahieren
	s.eax 		DMC_Time_RT.diff					//Ergebnis speicern
	l.ebx 		DMC_Time_RT.sum
	add.ebx 	eax								//Zur Summe addieren
	s.ebx 		DMC_Time_RT.sum					//Summe speichern
	l.ecx		  DMC_Time_RT.run
	inc 		  ecx								//Durchlaufzähler erhöhen
	s.ecx 		DMC_Time_RT.run					//Durchlaufzähler speichern
	cmp.eax		DMC_Time_RT._min					//mit Minimalzeit vergleichen
	jae			  LABEL_DMCcont
	s.eax 		DMC_Time_RT._min					//Minimalzeit speichern

LABEL_DMCcont
	cmp.eax 	DMC_Time_RT._max					//Mit Maximalzeit vergleichen
	jbe 		  LABEL_DMCcont1
	s.eax 		DMC_Time_RT._max					//Maximalzeit speichern

LABEL_DMCcont1
	l.eax		  ebx								//Summe in al laden
	imul.eax	eax,100							//*100 damit wir 2 Kommastellen haben
	x.edx 		edx
	idiv		  ecx								//durch Durchläufe dividieren
	s.eax		  DMC_Time_RT.avg					//Durchschnitt speichern
	popad

LABEL_DMCEND
	STI
#endif
//============================ Profiler end========================================================

END_FUNCTION
#endif

#pragma warning (disable:73)
FUNCTION VIRTUAL GLOBAL DiasMasterMain::I2CWriteOneByte
  VAR_INPUT
    AdressCDIAS		: UINT;
    pData		: ^USINT;
  END_VAR
  VAR_OUTPUT
    result		: DINT;
  END_VAR

	result:=-1;

END_FUNCTION

FUNCTION VIRTUAL GLOBAL DiasMasterMain::WriteEEData
  VAR_INPUT
    Adress		: UDINT;
    pData		: ^USINT;
    ui_length		: UINT;
    ui_offset		: UINT;
  END_VAR
  VAR_OUTPUT
    retval		: DINT;
  END_VAR

	retval:=-1;

END_FUNCTION
#pragma warning (default:73)
//[#ENGLISH]
//[>ui_value]value wich increases access time for ardware access
FUNCTION VIRTUAL GLOBAL DiasMasterMain::IncreaseHwAccessTime
  VAR_INPUT
    ui_value		: UINT;
  END_VAR

	ui_AddTime += ui_value;

END_FUNCTION

FUNCTION  DiasMasterMain::StartPll

	//start CDIAS Pll if available
	if ( p_CDIAS <> NIL ) then
		p_CDIAS^.us_Control.SyncOut	:= TRUE;
	end_if;

	//start DIAS Pll if available
	if ( p_DIAS <> NIL ) then
		p_DIAS^.us_Control.SyncOut	:= TRUE;
	end_if;

END_FUNCTION

FUNCTION DiasMasterMain::CorrectMyTaskTime

  //Only correct tasktime if we are Not connected with HwControl, we have a tasktime >1ms and PLL Trigger mode is correct
  if (ud_TaskTime > 1000) & ( CDIASSync <> NIL ) & ((CDIASSync + 2)^ AND 16#80) & HwControl = 0 then

    //set task time of DiasMaster to 1ms and select the right ms in RtWork
    if To_TaskObjectControl.ChangeObjectState( thispointer := this, actioncmd := 1, tasktype := OBJ_RT, debugobj := 0, newtime := 1 ) = 0 then
      b_TaskTimeCorrected := TRUE;
    else
      // failed to correct task time
    end_if;
  end_if;

END_FUNCTION

#ifdef _LSL_TARGETARCH_ARM
FUNCTION DiasMasterMain::LoadRtCyCode
  VAR
  	pIM   : ^USINT; // pointer to IM, where code should be stored
    pCode : ^USINT; // pointer on local memory, where code is stored
    i     : DINT;
  END_VAR

	// _IOSEGMENT    pointer to IM
	//	StartOfCode  load startoffset of programm in IM
	// #CodeRtCy     pointer on local memory, where code is stored
	// IPSub         maximum offset in local memory

  pIM := _IOSegment$^USINT + StartOfCode;
  pCode := #CodeRtCy[0];

  for i := 0 to (IPSub-1) do
    pIM^ := pCode^;

    pIM   += sizeof(USINT);
    pCode += sizeof(USINT);
  end_for;

END_FUNCTION
#else
FUNCTION AWL DiasMasterMain::LoadRtCyCode

	L.EDI		_IOSEGMENT   // pointer to IM
	L.EBX		StartOfCode  // load startoffset of programm in IM
	l.edx		#CodeRtCy    // pointer on local memory, where code is stored
	l.ecx		IPSub        // maximum offset in local memory
	inc			ecx          // increase by 1 to get length of used memory

LoadRtLoop
	l.al		(edx)
	s.al		(ebx+edi)
	inc			ebx
	inc			edx
	loop		LoadRtLoop

END_FUNCTION
#endif

FUNCTION VIRTUAL GLOBAL DiasMasterMain::GetObjectPath
	VAR_INPUT
		p_us_ObjectPath 	: ^USINT;
	END_VAR
	VAR_OUTPUT
		sd_retval 	: DINT;
	END_VAR

  if ( p_us_ObjectPath <> NIL ) then

    //set length of path = 1
    p_us_ObjectPath^ := 1;

#ifdef HWT_ucGetMyDomain
    if pHardwareTree then
      // at least CIL version 01.00.003 needed
      if pHardwareTree^.udVersion >= 16#1003 then
        // domain info byte
        ( p_us_ObjectPath + 1 )^ := HWT_ucGetMyDomain();
      else
        // domain info byte
        ( p_us_ObjectPath + 1 )^ := 0;
#ifdef HWC_LogError
        HWC_LogError(this, "@000E (DiasMasterMain::GetObjectPath) No domain info availbable: hardwaretree CIL version >= 01.00.003 needed");
#else
        TRACE("No domain info availbable: hardwaretree CIL version >= 01.00.003 needed");
#endif
      end_if;
    else
      // domain info byte
      ( p_us_ObjectPath + 1 )^ := 0;
    end_if;
#else
    // domain info byte
    ( p_us_ObjectPath + 1 )^ := 0;
#endif

    sd_retval := 0;

  else

    sd_retval := -1;

  end_if;

END_FUNCTION

FUNCTION VIRTUAL GLOBAL DiasMasterMain::SetObjectThisp
	VAR_INPUT
		p_us_ObjectPath 	: ^USINT;
		ud_thisp 	: UDINT;
	END_VAR
	VAR_OUTPUT
		sd_retval 	: DINT;
	END_VAR
  VAR
  	i : UINT;
    b_ModuleFound : BOOL;
  END_VAR

  if ( pHardwareTree <> NIL ) then

    sd_retval := HWT_ISETOBJECTTHISP(0,p_us_ObjectPath,ud_thisp);

  else

    sd_retval := 0;

  end_if;

  // Check if this pointer is already in the list
  b_ModuleFound := FALSE;
  if s_HWTModuleList.ui_Index then

    i := 0;
    repeat

      if (s_HWTModuleList.ap_ModuleList[i] = ud_thisp$pVirtualBase) then
        b_ModuleFound := TRUE;
      end_if;

      i += 1;
    until i >= s_HWTModuleList.ui_Index end_repeat;

  end_if;

  // Safe this pointer if it is not in the list
  if b_ModuleFound = FALSE &
     s_HWTModuleList.ui_Index < DIASMASTERC_MAX_MODULE_NO then
    s_HWTModuleList.ap_ModuleList[s_HWTModuleList.ui_Index] := ud_thisp$pVirtualBase;
    s_HWTModuleList.ui_Index += 1;
  end_if;

END_FUNCTION

FUNCTION VIRTUAL GLOBAL DiasMasterMain::GetObjectThisp
	VAR_INPUT
		p_us_ObjectPath 	: ^USINT;
	END_VAR
	VAR_OUTPUT
		ud_Thisp 	: UDINT;
	END_VAR

  if ( pHardwareTree <> NIL ) then

    ud_thisp := HWT_iGetObjectThisp(0,p_us_ObjectPath);

  else

    ud_thisp := 0;

  end_if;

END_FUNCTION

#ifdef _LSL_TARGETARCH_ARM
#pragma warning(disable:72 )
FUNCTION VIRTUAL GLOBAL DiasMasterMain::UpdateRtPostScan
  VAR
    pHandle  : ^OneHandle;
    i        : DINT;
  END_VAR
#pragma warning(default:72 )
#ifdef DM_DEBUG_ARM
  // This method is not supported with ARM
  ((0)$^USINT)^ := 0;
#endif

END_FUNCTION
#else

FUNCTION AWL VIRTUAL GLOBAL DiasMasterMain::UpdateRtPostScan

  // Function is called by HW-Control!

	l.ebx		  #HandlesRTPostScan
	lzxw.ecx	HandleNrRTPostScan
	jecxz		  NoRtProg

HandleLoopRt
	test.w		(ebx+OneHandle.Typ),DmCallProg
	jz			  NextHandleRt

	push		  ecx
	push		  ebx

	L.eax		  (ebx+OneHandle.thisp)
	LZXW.ECX	(ebx+OneHandle.Address)
	push		  ecx
	push		  eax

	call		  CallUpdataRtPostScan
	add.esp		8

	pop			  ebx
	pop			  ecx

NextHandleRt
	add.ebx		sizeof (OneHandle)
	loop		  HandleLoopRt

NoRtProg

END_FUNCTION
#endif

#ifdef _LSL_TARGETARCH_ARM
FUNCTION VIRTUAL GLOBAL DiasMasterMain::UpdateRtPostScan_IM
  VAR
    pHandle  : ^OneHandle;
    i        : UDINT;
  END_VAR

  // Function is called by HW-Control!
  if MasterON then
    // call update methods with thispointer
    if HandleNrRTPostScan then
      pHandle := #HandlesRTPostScan[0];

      for i := 0 to HandleNrRTPostScan-1 do
        if pHandle^.Typ AND DmCallProg then
          pHandle^.thisp^.UpdateRtPostScan(pHandle^.Address);
        end_if;

        pHandle += sizeof(OneHandle);
      end_for;
    end_if;

//LABEL_TimeSlice
    if (_IOSegment$^USINT + DmUserData + 4)^ then
      ud_ErrorCountTimeSliceStart += 1;
      if us_FirstTimeSliceStart = 0 then
        us_FirstTimeSliceStart := 1;
      end_if;
    end_if;
  end_if;

END_FUNCTION
#else

FUNCTION AWL VIRTUAL GLOBAL DiasMasterMain::UpdateRtPostScan_IM

  // Function is called by HW-Control!

  cmp.d     MasterON, 1
  jne       RT_End

	l.ebx		  #HandlesRTPostScan
	lzxw.ecx	HandleNrRTPostScan
	jecxz		  LABEL_TimeSlice

HandleLoopRt
	test.w		(ebx+OneHandle.Typ),DmCallProg
	jz			  NextHandleRt

	push		  ecx
	push		  ebx

	L.eax		  (ebx+OneHandle.thisp)
	LZXW.ECX	(ebx+OneHandle.Address)
	push		  ecx
	push		  eax

	call		  CallUpdataRtPostScan
	add.esp		8

	pop			  ebx
	pop			  ecx

NextHandleRt
	add.ebx		sizeof (OneHandle)
	loop		  HandleLoopRt

	//#SR010 start
LABEL_TimeSlice
  l.edi		  _IOSegment
	lzxb.eax	( edi + DmUserData + 4 )
	o.eax		  eax
	jz			  RT_end

	inc.d		  ud_ErrorCountTimeSliceStart
	cmp.b		  us_FirstTimeSliceStart,0
	jne			  RT_end
	l.b			  us_FirstTimeSliceStart,1
	//#SR010 end

RT_End

END_FUNCTION
#endif

FUNCTION DiasMasterMain::CallUpdataRtPostScan
	VAR_INPUT
		Thisp 	: pHwBase;
		Handle 	: UDINT;
	END_VAR

  thisp^.UpdateRtPostScan(handle);

END_FUNCTION

FUNCTION VIRTUAL GLOBAL DiasMasterMain::SetRetryCounterAvailability
	VAR_INPUT
		Port 	          : USINT;
		p_State 	      : ^IO_State;
		p_RetryCounter 	: ^DINT;
	END_VAR

  if s_RetryCounter.Quantity < 500 then
    s_RetryCounter.RetryCounter[s_RetryCounter.Quantity].Place          := Port;
    s_RetryCounter.RetryCounter[s_RetryCounter.Quantity].p_State        := p_State;
    s_RetryCounter.RetryCounter[s_RetryCounter.Quantity].p_RetryCounter := p_RetryCounter;
    s_RetryCounter.Quantity += 1;
  end_if;

END_FUNCTION

FUNCTION VIRTUAL DiasMasterMain::UpdateDIASRetryCounter
  VAR
    i                          : DINT;
    OldRetryCounter            : USINT;
    NewRetryCounter            : USINT;
    p_actualRetryCounterServer : ^UDINT;
    p_actualStateServer        : ^IO_State;
  END_VAR

  //get info how much DIAS moduls are connected
  i := s_RetryCounter.Quantity - 1 ;

  while i > - 1  do

    //load pointer to state server from counterstruct
    p_actualStateServer := (p_State + (i * sizeof(a_RetryStruct)))^$^IO_State;

    //check if pointer is valid
    if p_actualStateServer <> NIL then

      //check online state
      if MasterON then

        //compare if hw class state is ok
        if ((p_actualStateServer^$UINT) and 2#1100000000000011) = 0 then

          if DiasType = 2 then //check if we are intelligent master

            //load pointer to retrycounter server from counterstruct
            p_actualRetryCounterServer := (p_RetryCounter + (i * sizeof(a_RetryStruct)))^$^UDINT;

            //check if pointer is valid
            if p_actualRetryCounterServer <> NIL then

              //load retrycounter value from hardware
              NewRetryCounter := (p_ModuleRetryCnt$^USINT + (p_port + (i * sizeof(a_RetryStruct)))^)^;
              //get old value from counter
              OldRetryCounter := (p_OldRetryCounter + i)^;

              //check for differences
              if NewRetryCounter <> OldRetryCounter then

                //if new counter greater, no overflow ->
                if NewRetryCounter > OldRetryCounter then
                  p_actualRetryCounterServer^ += (NewRetryCounter - OldRetryCounter);
                else
                  //for overflow correction add 256
                  p_actualRetryCounterServer^ += (NewRetryCounter + 256 - OldRetryCounter);
                end_if;

                //set old counter to the value from new counter
                (p_OldRetryCounter + i)^ := NewRetryCounter;
              end_if;

            end_if;

          end_if;

        else

          //class state not ok, so set state pointer to nil - no more checks needed
          (p_State + (i * sizeof(a_RetryStruct)))^ := NIL;

        end_if;

      else
        //online state is 0, so signal error on class state server
        p_actualStateServer^$UINT := 16#FFFF;
      end_if;

    end_if;

    //decrement struct counter
    i -= 1;

  end_while;

END_FUNCTION

FUNCTION VIRTUAL GLOBAL DiasMasterMain::AddRequiredObject
	VAR_INPUT
		thisp 	: ^void;
	END_VAR

  if b_NotfirstCall = false then
    b_NotfirstCall := true;
    p_RequiredObjects := To_StdLib.Malloc(size:=(500*sizeof(^void)));
  end_if;

  if RequiredObjectCounter < 500 then
    (p_RequiredObjects + (RequiredObjectCounter * sizeof(^void)))^$^void := thisp;
    RequiredObjectCounter += 1;
  else
#ifdef HWC_LogError
    HWC_LogError(this, "@000F (DiasMasterMain::AddRequiredObject) Too many required object classes added");
#else
		TRACE( "DiasMaster: Too many required object classes added");
#endif
  end_if;

END_FUNCTION

#pragma warning(disable:137 )
FUNCTION VIRTUAL DiasMasterMain::CheckforRequiredError
  VAR
    i         : UINT;
    thisp     : ^virtualbase;
#ifndef HWC_LogError
    sz_name	  : array[ 0..255 ] of char;
#endif
    MyPara    : CmdStruct;
    MyResult  : results;
    DiasError : BOOL;
    CdiasError: BOOL;
  END_VAR

  if RequiredObjectCounter > 0 then
    //--- init the newInst command
    MyPara.uiCmd := DM_CHECK_REQUIRED_ERROR;
    CdiasError  := false;
    DiasError   := false;
    for i := 0 to (RequiredObjectCounter -1) do
      thisp := (p_RequiredObjects + (i * sizeof(^void)))^$^virtualbase;
      //--- init result for next call
      MyResult.aData[0] := 16#FF;
      MyResult.aData[1] := 16#FF;
      if (thisp^.NewInst(#MyPara, #MyResult) = ERROR) then
        //Required Error!

        if (MyResult.aData[1] = CDIAS_MODULE) then
          CdiasError := true;
        end_if;
        if (MyResult.aData[1] = DIAS_MODULE) then
          DiasError := true;
        end_if;

#ifdef HWC_LogError
        HWC_LogError(thisp, "@0010 (DiasMasterMain::CheckforRequiredError) Required Error triggerd by this object");
#else
        _GetObjName( thisp, #sz_name[ 0 ] );
        if RequiredErrors = 0 then
          Trace ("DiasMaster: Required Error triggerd by object(s):");
        end_if;
        Trace (#sz_name[ 0 ] );
#endif

        RequiredErrors +=1;
      end_if;
    end_for;

    if RequiredErrors > 0 then

      if ( IsClientConnected( #To_HwControl ) ) then
        To_HwControl.Write(0);
      end_if;

      case _WhoAmI of
        DESTPLC_WINPC_98,    // LARS, Standard PC, Win98/ME
        DESTPLC_WINPC_NT,    // LARS, Standard PC, WinNT/Win2000/WinXP
        DESTPLC_WINIPC_98,   // LARS, IPC, Win98/ME
        DESTPLC_WINIPC_NT:   // LARS, IPC, WinNT/Win2000/WinXP

          //LARS
          //RamAnd: Don't execute a required error when target platform is lars due to SA 40955

      else
        //--- rtk-os
          if (_rtosversion >= 16#12DC) & (CdiasError = true)then   // _rtosversion >= 1.2.220
            To_OSKernel.AddToServiceProvider(command:="exec climsg 70 A CDIAS module is set required, but there is no CDIAS Module", immediatly:=1);  //stop application
          elsif (_rtosversion >= 16#12DC) & (DiasError = true) then // _rtosversion >= 1.2.220
            To_OSKernel.AddToServiceProvider(command:="exec climsg 25 A DIAS module is set required, but there is no DIAS Module", immediatly:=1);  //stop application
          else
            To_OSKernel.Reset();  //stop application, because this OS doesn't support the message and the CPU state
          end_if;
      end_case;

    end_if;

    To_StdLib.Free(p_RequiredObjects);

  end_if;

END_FUNCTION
#pragma warning(Default:137 )

FUNCTION VIRTUAL GLOBAL DiasMasterMain::SetRequiredError
	VAR_INPUT
		p_this 	: ^HWBase;
	END_VAR
#ifndef HWC_LogError
  VAR
 		sz_name	: array[ 0..255 ] of char;
  END_VAR
#endif

  //Required Error!

  //log the object responsable
#ifdef HWC_LogError
  HWC_LogError(p_this, "@0011 (DiasMasterMain::SetRequiredError) Required Error triggerd by this object");
#else
  _GetObjName( p_this, #sz_name[ 0 ] );
  if RequiredErrors = 0 then
    Trace ("Required Error triggerd by object(s):");
  end_if;
  Trace (#sz_name[ 0 ] );
#endif

  RequiredErrors +=1;

  if RequiredErrors > 0 then

    if ( IsClientConnected( #To_HwControl ) ) then
      To_HwControl.Write(0);
    end_if;

    MasterON := 0;
    To_OSKernel.Reset();

  end_if;

END_FUNCTION

FUNCTION DiasMasterMain::CallSafetyManager

  SafetyManagerThis^.CyWork(0);

END_FUNCTION

FUNCTION VIRTUAL GLOBAL DiasMasterMain::Control::NewInst
	VAR_INPUT
		pPara 	: ^CmdStruct;
		pResult 	: ^Results;
	END_VAR
	VAR_OUTPUT
		ret_code 	: IprStates;
	END_VAR
  VAR
  	ui_CurrentHandleNr : UINT;
    // local variables for the Requested HWTString
    pStr_HWTRequested     : ^CHAR;
    b_ModuleFound : BOOL;
  END_VAR

  ui_CurrentHandleNr  := 0;
  // local variables for the Requested HWTString
  pStr_HWTRequested   := NIL;
  b_ModuleFound       := FALSE;

  ret_code := ERROR;

  CASE pPara^.uiCmd OF
    //**********************************************************************************************************************************************************
    CMD_GET_HARDWARE_TREE_ENTRY:

      //Set Errors
      pResult^.aData[0]$t_HWCGetHardwareTreeEntryOut.retcode := _HWC_RETVAL_ERROR;
      ret_code := ERROR;

      pStr_HWTRequested     := pPara^.aPara[0]$t_HWCGetHardwareDiagnosisIn.pStr_HardewareTreeEntry;

      //First HWT Path
      if pStr_HWTRequested = nil then

        //DiasMaster always has the same object path, store it on the variable
        ud_DiasMasterPosition := DIASMASTERC_OBJECT_PATH_CDIAS;

        ret_code := READY;
        pResult^.aData$t_HWCGetHardwareTreeEntryOut.retcode := _HWC_RETVAL_OK_HWTSTR_RETURNED;
        pResult^.aData[0]$t_HWCGetHardwareTreeEntryOut.pStr_NextHardewareTreeEntry := (#ud_DiasMasterPosition)$^CHAR;

      //Only possible for Diasmaster own HWT Path
      elsif (pStr_HWTRequested^$USINT = 2) & (pStr_HWTRequested^$UDINT = DIASMASTERC_OBJECT_PATH_CDIAS) then

        //DiasMaster always has the same object path, store it on the variable
        ud_DiasMasterPosition := DIASMASTERC_OBJECT_PATH_DIAS;

        ret_code := READY;
        pResult^.aData$t_HWCGetHardwareTreeEntryOut.retcode := _HWC_RETVAL_OK_HWTSTR_RETURNED;
        pResult^.aData[0]$t_HWCGetHardwareTreeEntryOut.pStr_NextHardewareTreeEntry := (#ud_DiasMasterPosition)$^CHAR;

      elsif (pStr_HWTRequested^$USINT = 2) & (pStr_HWTRequested^$UDINT = DIASMASTERC_OBJECT_PATH_DIAS) then

        // Check i list is valid
        if s_HWTModuleList.ui_Index > 0 then

          // Call 1st entry in list
          if s_HWTModuleList.ap_ModuleList[0] then
            ret_code := s_HWTModuleList.ap_ModuleList[0]^.NewInst(pPara:=pPara, pResult:=pResult);
          end_if;
        else
          // Dias/CDIAS Master found, but no modules connected.
          ret_code := READY;
          pResult^.aData[0]$t_HWCGetHardwareTreeEntryOut.retcode := _HWC_RETVAL_OK_MODULE_FOUND;
        end_if;

      else

        // Only Error case is returned from the newInst
        ret_code := READY;
        pResult^.aData[0]$t_HWCGetHardwareTreeEntryOut.retcode := _HWC_RETVAL_OK_MODULE_FOUND;

        // Search for module with passed HWT string
        if s_HWTModuleList.ui_Index > 0 &
           s_HWTModuleList.ui_Index <= DIASMASTERC_MAX_MODULE_NO then

          ui_CurrentHandleNr := 0;
          b_ModuleFound := FALSE;

          repeat

            // Search for the passed HWT-Strubg
            if s_HWTModuleList.ap_ModuleList[ui_CurrentHandleNr] then
              ret_code := s_HWTModuleList.ap_ModuleList[ui_CurrentHandleNr]^.NewInst(pPara:=pPara, pResult:=pResult);
            end_if;

            ui_CurrentHandleNr += 1;

            if ret_code = READY & pResult^.aData$t_HWCGetHardwareTreeEntryOut.retcode = _HWC_RETVAL_OK_MODULE_FOUND then
              // If Module was found
              b_ModuleFound := TRUE;
              exit;

            end_if;

          until ui_CurrentHandleNr >= s_HWTModuleList.ui_Index end_repeat;

          if b_ModuleFound &                                    // Module was found
             ui_CurrentHandleNr < s_HWTModuleList.ui_Index then // and the next entry is in the list

            repeat

              // Call next valid Module
              if s_HWTModuleList.ap_ModuleList[ui_CurrentHandleNr] then
                ret_code := s_HWTModuleList.ap_ModuleList[ui_CurrentHandleNr]^.NewInst(pPara:=pPara, pResult:=pResult);
                return;
              end_if;

            until ui_CurrentHandleNr >= s_HWTModuleList.ui_Index end_repeat;

            // Already set
//          else
//            // Dias/CDIAS Module found, but no further modules connected.
//            ret_code := READY;
//            pResult^.aData[0]$t_HWCGetHardwareTreeEntryOut.retcode := _HWC_RETVAL_OK_MODULE_FOUND;
          end_if;

          // Already set
//        else
//          // Dias/CDIAS Master found, but no modules connected.
//          ret_code := READY;
//          pResult^.aData[0]$t_HWCGetHardwareTreeEntryOut.retcode := _HWC_RETVAL_OK_MODULE_FOUND;
        end_if;
      end_if;

    //**********************************************************************************************************************************************************
    CMD_GET_HARDWARE_DIAGNOSIS:

      //Set Errors
      pResult^.aData[0]$t_HWCGetHardwareTreeEntryOut.retcode := _HWC_RETVAL_ERROR;
      ret_code := ERROR;

      pStr_HWTRequested     := pPara^.aPara[0]$t_HWCGetHardwareDiagnosisIn.pStr_HardewareTreeEntry;

      if pStr_HWTRequested$^UINT^ > 2 then

        // Search for module with passed HWT string
        if s_HWTModuleList.ui_Index > 0 &
           s_HWTModuleList.ui_Index <= DIASMASTERC_MAX_MODULE_NO then

          // Change Command to CMD_GET_HARDWARE_TREE_ENTRY search for the module
          pPara^.uiCmd := CMD_GET_HARDWARE_TREE_ENTRY;

          ui_CurrentHandleNr := 0;
          repeat

            ret_code := s_HWTModuleList.ap_ModuleList[ui_CurrentHandleNr]^.NewInst(pPara:=pPara, pResult:=pResult);

            if ret_code = READY & pResult^.aData$t_HWCGetHardwareTreeEntryOut.retcode = _HWC_RETVAL_OK_MODULE_FOUND then

              // Get Diagnosis of Module just found
              pPara^.uiCmd := CMD_GET_HARDWARE_DIAGNOSIS;

              ret_code := s_HWTModuleList.ap_ModuleList[ui_CurrentHandleNr]^.NewInst(pPara:=pPara, pResult:=pResult);

              return;
            end_if;

            ui_CurrentHandleNr += 1;

          until ui_CurrentHandleNr >= s_HWTModuleList.ui_Index end_repeat;

        end_if;

      // Check for diasmaster
      elsif (pStr_HWTRequested^$USINT = 2) &
         (pStr_HWTRequested^$UDINT = DIASMASTERC_OBJECT_PATH_CDIAS | pStr_HWTRequested^$UDINT = DIASMASTERC_OBJECT_PATH_DIAS ) then

        pResult^.aData$t_HWCGetHardwareDiagnosisOut.retcode     := _HWC_RETVAL_OK;
        ret_code := READY;
      end_if;
//**********************************************************************************************************************************************************
    CMD_HWC_ERROR_TO_DIASM:
      // we need to stop the cyclic (rt is stopped, since it's no longer called by the hw control object)
      MasterOn := 0;
      ImOff := 1;
      SkipCy := true;

//**********************************************************************************************************************************************************
    CMD_SET_POSTINIT_DONE:
      ret_code := READY;
      b_IsPostInitDone := TRUE;

//**********************************************************************************************************************************************************
    CMD_IS_POSTINIT_DONE:

      ret_code := READY;
      pResult^.uiLng    := sizeof(BOOL);
      pResult^.aData[0]$BOOL := b_IsPostInitDone;

//**********************************************************************************************************************************************************
    else

      ret_code := DiasMaster::Control.NewInst(pPara, pResult);

  END_CASE;

END_FUNCTION
